// ---- SelfTests/TestCases/TestSuite_EventDelivery/Test_EventDeleteLostSequence.TcPOU
{region 'Documentation'}
(*!
<summary>Verifies deletion progress stops at retained events when the requested sequence was lost.</summary>
<description>
Four primary events plus the capacity diagnostic fill five usable slots. Publications 6
and 7 fail, creating a real sequence gap. Request 6 exhausts the retained prefix at 5 and
appends diagnostic 8. Request 7 must leave that newer head intact and append diagnostic 9.
No sequence, FIFO index or private subject field is modified to arrange these cases.
The real subject binds only local storage; expected findings remain in that storage.
Checking Assertions retain the outer selftest publisher. Each run reinitializes the subject.
</description>
*)
{endregion}
FUNCTION_BLOCK Test_EventDeleteLostSequence EXTENDS TestCaseBase
VAR
    FSubject : EventBuffer;
    FEvents : ARRAY[1..BufferLength] OF ST_Event;
    FFifo : ST_FifoStatus;
    FBufferStatus : ST_EventBufferStatus;
    FPerformed : BOOL;
    FChecked : BOOL;
    FLostTargets : AssertTrue;
    FLostTargetsMatches : BOOL;
    FActualProgress : AssertTrue;
    FActualProgressMatches : BOOL;
    FExhaustionDiagnostic : AssertTrue;
    FExhaustionDiagnosticMatches : BOOL;
    FNewerHeadPreserved : AssertTrue;
    FNewerHeadPreservedMatches : BOOL;
    FGapDiagnostic : AssertTrue;
    FGapDiagnosticMatches : BOOL;
END_VAR
VAR CONSTANT
    BufferLength : UINT := 6;
END_VAR

SUPER^();

{region 'Documentation'}
(*!
<summary>Contributes each checking Assertion once.</summary>
*)
{endregion}
METHOD PROTECTED AggregateResults
VAR_INPUT
    Aggregator : I_ResultAggregator; //! Borrowed result sink owned by the outer Test Case; add this test's checking Assertions without resetting or retaining the sink.
END_VAR
Aggregator.AddProvider(Provider := FLostTargets);
Aggregator.AddProvider(Provider := FActualProgress);
Aggregator.AddProvider(Provider := FExhaustionDiagnostic);
Aggregator.AddProvider(Provider := FNewerHeadPreserved);
Aggregator.AddProvider(Provider := FGapDiagnostic);
END_METHOD

{region 'Documentation'}
(*!
<summary>Requires all checking Assertions to be initialized.</summary>
*)
{endregion}
METHOD PROTECTED CheckInitialization : BOOL //! TRUE when the inherited initialization check and this concrete fixture check both accept the setup.
CheckInitialization := FALSE;
IF NOT SUPER^.CheckInitialization() THEN
    RETURN;
END_IF;

CheckInitialization := FLostTargets.IsInitialized
    AND FActualProgress.IsInitialized
    AND FExhaustionDiagnostic.IsInitialized
    AND FNewerHeadPreserved.IsInitialized
    AND FGapDiagnostic.IsInitialized;
END_METHOD

{region 'Documentation'}
(*!
<summary>Initializes the checking Assertions for one test state.</summary>
*)
{endregion}
METHOD PROTECTED Configure
FPreparationStateCount := 0;
FTestStateCount := 1;
FLostTargets.Initialize(Parent := THIS^,
    AssertionName := 'LostTargets');
FActualProgress.Initialize(Parent := THIS^,
    AssertionName := 'ActualProgress');
FExhaustionDiagnostic.Initialize(Parent := THIS^,
    AssertionName := 'ExhaustionDiagnostic');
FNewerHeadPreserved.Initialize(Parent := THIS^,
    AssertionName := 'NewerHeadPreserved');
FGapDiagnostic.Initialize(Parent := THIS^,
    AssertionName := 'GapDiagnostic');
END_METHOD

{region 'Documentation'}
(*!
<summary>Fills the buffer and verifies that sequences 6 and 7 were assigned but not retained.</summary>
*)
{endregion}
METHOD PRIVATE CreateLostTargets
VAR
    Index : UINT;
    WriteResult : INT;
END_VAR
FLostTargetsMatches := TRUE;
FOR Index := 1 TO 4 DO
    WriteResult := FSubject.PublishEvent(Event := CreateFrameworkEvent(Name := 'LocalGap',
        State := E_State.Running,
        Severity := E_EventSeverity.Info,
        Message := UINT_TO_STRING(Index)));
    FLostTargetsMatches := FLostTargetsMatches AND (WriteResult = UINT_TO_INT(Index));
END_FOR;
FOR Index := 6 TO 7 DO
    WriteResult := FSubject.PublishEvent(Event := CreateFrameworkEvent(Name := 'Lost',
        State := E_State.Running,
        Severity := E_EventSeverity.Info,
        Message := UINT_TO_STRING(Index)));
    FLostTargetsMatches := FLostTargetsMatches AND (WriteResult = TO_INT(E_FifoResult.NoTransfer));
END_FOR;
FLostTargetsMatches := FLostTargetsMatches AND FFifo.BufferFull
    AND (FFifo.ElementCount = 5) AND (FFifo.IndexOut = 1) AND (FFifo.IndexIn = 6)
    AND (FBufferStatus.SequenceId = 7) AND (FBufferStatus.DeletedSequenceId = 0)
    AND (FBufferStatus.LostEventCount = 2);
FOR Index := 1 TO 5 DO
    FLostTargetsMatches := FLostTargetsMatches AND (FEvents[Index].SequenceId = UINT_TO_UDINT(Index));
END_FOR;
END_METHOD

{region 'Documentation'}
(*!
<summary>A lost target below the current head must not delete that newer event or advance the watermark.</summary>
*)
{endregion}
METHOD PRIVATE DeleteBeforeNewerHead
VAR
    Request : UDINT;
    HeadBeforeRequest : ST_Event;
END_VAR
HeadBeforeRequest := FEvents[6];
Request := 7;
FSubject.ProcessDeleteRequest(SequenceId := Request);
FNewerHeadPreservedMatches := (Request = 0) AND (FBufferStatus.DeletedSequenceId = 5)
    AND (FBufferStatus.LostEventCount = 2)
    AND (FFifo.IndexOut = 6) AND (FFifo.IndexIn = 2) AND (FFifo.ElementCount = 2)
    AND (FEvents[6].SequenceId = 8)
    AND (FEvents[6].SequenceId = HeadBeforeRequest.SequenceId)
    AND (FEvents[6].Timestamp = HeadBeforeRequest.Timestamp)
    AND (FEvents[6].OwnerScope = HeadBeforeRequest.OwnerScope)
    AND (FEvents[6].EventType = HeadBeforeRequest.EventType)
    AND (FEvents[6].Severity = HeadBeforeRequest.Severity)
    AND (FEvents[6].Name = HeadBeforeRequest.Name)
    AND (FEvents[6].ResourceName = HeadBeforeRequest.ResourceName)
    AND (FEvents[6].State = HeadBeforeRequest.State)
    AND (FEvents[6].Result = HeadBeforeRequest.Result)
    AND (FEvents[6].Message = HeadBeforeRequest.Message);
FGapDiagnosticMatches := (FBufferStatus.SequenceId = 9)
    AND (FEvents[1].SequenceId = 9) AND (FEvents[1].OwnerScope = E_OwnerScope.Framework)
    AND (FEvents[1].EventType = E_EventType.Framework)
    AND (FEvents[1].Severity = E_EventSeverity.Warning) AND (FEvents[1].Name = 'EventBuffer');
END_METHOD

{region 'Documentation'}
(*!
<summary>Deletion exhausts at sequence 5; the newly appended diagnostic is not part of that prefix.</summary>
*)
{endregion}
METHOD PRIVATE DeleteBeyondRetainedTail
VAR
    Request : UDINT;
    Index : UINT;
END_VAR
Request := 6;
FSubject.ProcessDeleteRequest(SequenceId := Request);
FActualProgressMatches := (Request = 0) AND (FBufferStatus.DeletedSequenceId = 5)
    AND (FBufferStatus.LostEventCount = 2);
FOR Index := 1 TO 5 DO
    FActualProgressMatches := FActualProgressMatches AND (FEvents[Index].SequenceId = 0)
        AND (FEvents[Index].Timestamp = 0) AND (FEvents[Index].Name = '') AND (FEvents[Index].Message = '');
END_FOR;
FExhaustionDiagnosticMatches := (FBufferStatus.SequenceId = 8)
    AND NOT FFifo.BufferEmpty AND (FFifo.ElementCount = 1)
    AND (FFifo.IndexOut = 6) AND (FFifo.IndexIn = 1)
    AND (FEvents[6].SequenceId = 8) AND (FEvents[6].OwnerScope = E_OwnerScope.Framework)
    AND (FEvents[6].EventType = E_EventType.Framework)
    AND (FEvents[6].Severity = E_EventSeverity.Warning) AND (FEvents[6].Name = 'EventBuffer');
END_METHOD

{region 'Documentation'}
(*!
<summary>Creates two lost targets through overflow, then exercises exhaustion and a newer FIFO head.</summary>
*)
{endregion}
METHOD PRIVATE ExerciseBuffer
IF NOT FSubject.Initialize(Buffer := FEvents,
    FifoControl := FFifo,
    Status := FBufferStatus) THEN
    Error(Message := 'Local Event Buffer initialization failed.');
    RETURN;
END_IF;

CreateLostTargets();
DeleteBeyondRetainedTail();
DeleteBeforeNewerHead();
END_METHOD

{region 'Documentation'}
(*!
<summary>Completes abort without asynchronous work.</summary>
*)
{endregion}
METHOD PROTECTED ProcessAbort
VAR_INPUT
    Enable : BOOL; //! Phase permission supplied by the owning Test Case; FALSE does not authorize progression, while observation may continue.
END_VAR
IF Enable THEN
    CompleteAbort();
END_IF;
END_METHOD

{region 'Documentation'}
(*!
<summary>Evaluates captured observations after the scenario has finished.</summary>
*)
{endregion}
METHOD PROTECTED ProcessAssertions
VAR_INPUT
    Enable : BOOL; //! Phase permission supplied by the owning Test Case; FALSE does not authorize progression, while observation may continue.
END_VAR
VAR
    Evaluate : BOOL;
END_VAR
Evaluate := Enable AND FPerformed;
FLostTargets(Enable := Evaluate,
    State := State,
    IN := FLostTargetsMatches);
FActualProgress(Enable := Evaluate,
    State := State,
    IN := FActualProgressMatches);
FExhaustionDiagnostic(Enable := Evaluate,
    State := State,
    IN := FExhaustionDiagnosticMatches);
FNewerHeadPreserved(Enable := Evaluate,
    State := State,
    IN := FNewerHeadPreservedMatches);
FGapDiagnostic(Enable := Evaluate,
    State := State,
    IN := FGapDiagnosticMatches);
IF Evaluate THEN
    FChecked := TRUE;
END_IF;
END_METHOD

{region 'Documentation'}
(*!
<summary>No Preparation phase is needed.</summary>
*)
{endregion}
METHOD PROTECTED ProcessPreparations
VAR_INPUT
    // SA0033: Required override without Preparation work.
    {attribute 'analysis' := '-33'}
    Enable : BOOL; //! Phase permission supplied by the owning Test Case; FALSE does not authorize progression, while observation may continue.
END_VAR
END_METHOD

{region 'Documentation'}
(*!
<summary>Resets observations and schedules a fresh subject initialization.</summary>
*)
{endregion}
METHOD PROTECTED ProcessReset
FPerformed := FALSE;
FChecked := FALSE;
FLostTargets.Reset();
FLostTargetsMatches := FALSE;
FActualProgress.Reset();
FActualProgressMatches := FALSE;
FExhaustionDiagnostic.Reset();
FExhaustionDiagnosticMatches := FALSE;
FNewerHeadPreserved.Reset();
FNewerHeadPreservedMatches := FALSE;
FGapDiagnostic.Reset();
FGapDiagnosticMatches := FALSE;
CompleteReset();
END_METHOD

{region 'Documentation'}
(*!
<summary>Runs the bounded scenario once before Assertion evaluation.</summary>
*)
{endregion}
METHOD PROTECTED ProcessTests
VAR_INPUT
    Enable : BOOL; //! Phase permission supplied by the owning Test Case; FALSE does not authorize progression, while observation may continue.
END_VAR
IF NOT Enable THEN
    RETURN;
END_IF;
IF FChecked THEN
    CompleteTests();
    RETURN;
END_IF;

IF NOT FPerformed THEN
    ExerciseBuffer();
    FPerformed := TRUE;
END_IF;
END_METHOD

END_FUNCTION_BLOCK

// ---- SelfTests/TestCases/TestSuite_EventDelivery/Test_EventDeleteCommandBoundary.TcPOU
{region 'Documentation'}
(*!
<summary>Verifies DeleteSequenceId consumption at explicit call boundaries across successive PLC cycles.</summary>
<description>
Uses the actual field of a local ST_EventBufferCommand as VAR_IN_OUT, not a copied request.
A higher watermark replaces an earlier value before the call. Another is queued after return,
survives publication in the next cycle and is consumed only by the following delete call.
Zero after successful or rejected processing must not replay deletion or diagnostics.
No write occurs inside ProcessDeleteRequest: this scenario does not exercise its changed-value
branch or establish atomicity against ADS writes between comparison and clearing.
The real subject binds only local storage; expected findings remain in that storage.
Checking Assertions retain the outer selftest publisher. Each run reinitializes the subject.
</description>
*)
{endregion}
FUNCTION_BLOCK Test_EventDeleteCommandBoundary EXTENDS TestCaseBase
VAR
    FSubject : EventBuffer;
    FEvents : ARRAY[1..BufferLength] OF ST_Event;
    FFifo : ST_FifoStatus;
    FBufferStatus : ST_EventBufferStatus;
    FPerformed : BOOL;
    FChecked : BOOL;
    FCommands : ST_EventBufferCommand;
    FStep : UINT;
    FBeforeCall : AssertTrue;
    FBeforeCallMatches : BOOL;
    FPending : AssertTrue;
    FPendingMatches : BOOL;
    FNextCall : AssertTrue;
    FNextCallMatches : BOOL;
    FZeroNoReplay : AssertTrue;
    FZeroNoReplayMatches : BOOL;
    FRejectedNoReplay : AssertTrue;
    FRejectedNoReplayMatches : BOOL;
END_VAR
VAR CONSTANT
    BufferLength : UINT := 10;
    Arrange : UINT := 0;
    ReplaceBeforeCall : UINT := 1;
    ObservePending : UINT := 2;
    ConsumePending : UINT := 3;
    ObserveCleared : UINT := 4;
    RejectFuture : UINT := 5;
    ObserveRejected : UINT := 6;
END_VAR

SUPER^();

{region 'Documentation'}
(*!
<summary>Contributes each checking Assertion once.</summary>
*)
{endregion}
METHOD PROTECTED AggregateResults
VAR_INPUT
    Aggregator : I_ResultAggregator; //! Borrowed result sink owned by the outer Test Case; add this test's checking Assertions without resetting or retaining the sink.
END_VAR
Aggregator.AddProvider(Provider := FBeforeCall);
Aggregator.AddProvider(Provider := FPending);
Aggregator.AddProvider(Provider := FNextCall);
Aggregator.AddProvider(Provider := FZeroNoReplay);
Aggregator.AddProvider(Provider := FRejectedNoReplay);
END_METHOD

{region 'Documentation'}
(*!
<summary>Requires all checking Assertions to be initialized.</summary>
*)
{endregion}
METHOD PROTECTED CheckInitialization : BOOL //! TRUE when the inherited initialization check and this concrete fixture check both accept the setup.
CheckInitialization := FALSE;
IF NOT SUPER^.CheckInitialization() THEN
    RETURN;
END_IF;

CheckInitialization := FBeforeCall.IsInitialized
    AND FPending.IsInitialized
    AND FNextCall.IsInitialized
    AND FZeroNoReplay.IsInitialized
    AND FRejectedNoReplay.IsInitialized;
END_METHOD

{region 'Documentation'}
(*!
<summary>Initializes the checking Assertions for one test state.</summary>
*)
{endregion}
METHOD PROTECTED Configure
FPreparationStateCount := 0;
FTestStateCount := 1;
FBeforeCall.Initialize(Parent := THIS^,
    AssertionName := 'BeforeCall');
FPending.Initialize(Parent := THIS^,
    AssertionName := 'Pending');
FNextCall.Initialize(Parent := THIS^,
    AssertionName := 'NextCall');
FZeroNoReplay.Initialize(Parent := THIS^,
    AssertionName := 'ZeroNoReplay');
FRejectedNoReplay.Initialize(Parent := THIS^,
    AssertionName := 'RejectedNoReplay');
END_METHOD

{region 'Documentation'}
(*!
<summary>Completes abort without asynchronous work.</summary>
*)
{endregion}
METHOD PROTECTED ProcessAbort
VAR_INPUT
    Enable : BOOL; //! Phase permission supplied by the owning Test Case; FALSE does not authorize progression, while observation may continue.
END_VAR
IF Enable THEN
    CompleteAbort();
END_IF;
END_METHOD

{region 'Documentation'}
(*!
<summary>Evaluates captured observations after the scenario has finished.</summary>
*)
{endregion}
METHOD PROTECTED ProcessAssertions
VAR_INPUT
    Enable : BOOL; //! Phase permission supplied by the owning Test Case; FALSE does not authorize progression, while observation may continue.
END_VAR
VAR
    Evaluate : BOOL;
END_VAR
Evaluate := Enable AND FPerformed;
FBeforeCall(Enable := Evaluate,
    State := State,
    IN := FBeforeCallMatches);
FPending(Enable := Evaluate,
    State := State,
    IN := FPendingMatches);
FNextCall(Enable := Evaluate,
    State := State,
    IN := FNextCallMatches);
FZeroNoReplay(Enable := Evaluate,
    State := State,
    IN := FZeroNoReplayMatches);
FRejectedNoReplay(Enable := Evaluate,
    State := State,
    IN := FRejectedNoReplayMatches);
IF Evaluate THEN
    FChecked := TRUE;
END_IF;
END_METHOD

{region 'Documentation'}
(*!
<summary>No Preparation phase is needed.</summary>
*)
{endregion}
METHOD PROTECTED ProcessPreparations
VAR_INPUT
    // SA0033: Required override without Preparation work.
    {attribute 'analysis' := '-33'}
    Enable : BOOL; //! Phase permission supplied by the owning Test Case; FALSE does not authorize progression, while observation may continue.
END_VAR
END_METHOD

{region 'Documentation'}
(*!
<summary>Resets observations and schedules a fresh subject initialization.</summary>
*)
{endregion}
METHOD PROTECTED ProcessReset
FPerformed := FALSE;
FChecked := FALSE;
FStep := Arrange;
FCommands.Reset := FALSE;
FCommands.DeleteSequenceId := 0;
FBeforeCall.Reset();
FBeforeCallMatches := FALSE;
FPending.Reset();
FPendingMatches := FALSE;
FNextCall.Reset();
FNextCallMatches := FALSE;
FZeroNoReplay.Reset();
FZeroNoReplayMatches := FALSE;
FRejectedNoReplay.Reset();
FRejectedNoReplayMatches := FALSE;
CompleteReset();
END_METHOD

{region 'Documentation'}
(*!
<summary>Advances the scenario until its final observation has been evaluated.</summary>
*)
{endregion}
METHOD PROTECTED ProcessTests
VAR_INPUT
    Enable : BOOL; //! Phase permission supplied by the owning Test Case; FALSE does not authorize progression, while observation may continue.
END_VAR
IF NOT Enable THEN
    RETURN;
END_IF;
IF FChecked THEN
    CompleteTests();
    RETURN;
END_IF;

IF NOT FPerformed THEN
    StateMachine();
END_IF;
END_METHOD

{region 'Documentation'}
(*!
<summary>Advances one boundary scenario step per enabled test cycle.</summary>
*)
{endregion}
METHOD PRIVATE StateMachine
VAR
    Index : UINT;
    WriteResult : INT;
END_VAR
CASE FStep OF
    Arrange:
        IF NOT FSubject.Initialize(Buffer := FEvents,
            FifoControl := FFifo,
            Status := FBufferStatus) THEN
            Error(Message := 'Local Event Buffer initialization failed.');
            RETURN;
        END_IF;
        FBeforeCallMatches := TRUE;
        FOR Index := 1 TO 4 DO
            WriteResult := FSubject.PublishEvent(Event := CreateFrameworkEvent(Name := 'LocalCommand',
                State := E_State.Running,
                Severity := E_EventSeverity.Info,
                Message := UINT_TO_STRING(Index)));
            FBeforeCallMatches := FBeforeCallMatches AND (WriteResult = UINT_TO_INT(Index));
        END_FOR;
        FStep := ReplaceBeforeCall;

    ReplaceBeforeCall:
        FCommands.DeleteSequenceId := 1;
        FCommands.DeleteSequenceId := 2;
        FSubject.ProcessDeleteRequest(SequenceId := FCommands.DeleteSequenceId);
        FBeforeCallMatches := FBeforeCallMatches AND (FCommands.DeleteSequenceId = 0)
            AND (FBufferStatus.DeletedSequenceId = 2) AND (FBufferStatus.SequenceId = 4)
            AND (FFifo.IndexOut = 3) AND (FFifo.IndexIn = 5) AND (FFifo.ElementCount = 2)
            AND (FEvents[1].SequenceId = 0) AND (FEvents[2].SequenceId = 0)
            AND (FEvents[3].SequenceId = 3) AND (FEvents[4].SequenceId = 4);
        FCommands.DeleteSequenceId := 4;
        FStep := ObservePending;

    ObservePending:
        WriteResult := FSubject.PublishEvent(Event := CreateFrameworkEvent(Name := 'LocalCommand',
            State := E_State.Running,
            Severity := E_EventSeverity.Info,
            Message := 'Published while deletion is pending.'));
        FPendingMatches := (WriteResult = 5) AND (FCommands.DeleteSequenceId = 4)
            AND (FBufferStatus.DeletedSequenceId = 2) AND (FBufferStatus.SequenceId = 5)
            AND (FFifo.IndexOut = 3) AND (FFifo.IndexIn = 6) AND (FFifo.ElementCount = 3)
            AND (FEvents[3].SequenceId = 3) AND (FEvents[4].SequenceId = 4)
            AND (FEvents[5].SequenceId = 5);
        FStep := ConsumePending;

    ConsumePending:
        FSubject.ProcessDeleteRequest(SequenceId := FCommands.DeleteSequenceId);
        FNextCallMatches := (FCommands.DeleteSequenceId = 0)
            AND (FBufferStatus.DeletedSequenceId = 4) AND (FBufferStatus.SequenceId = 5)
            AND (FFifo.IndexOut = 5) AND (FFifo.IndexIn = 6) AND (FFifo.ElementCount = 1)
            AND (FEvents[3].SequenceId = 0) AND (FEvents[4].SequenceId = 0)
            AND (FEvents[5].SequenceId = 5);
        FStep := ObserveCleared;

    ObserveCleared:
        FSubject.ProcessDeleteRequest(SequenceId := FCommands.DeleteSequenceId);
        FZeroNoReplayMatches := (FCommands.DeleteSequenceId = 0)
            AND (FBufferStatus.DeletedSequenceId = 4) AND (FBufferStatus.SequenceId = 5)
            AND (FFifo.IndexOut = 5) AND (FFifo.IndexIn = 6) AND (FFifo.ElementCount = 1)
            AND (FEvents[5].SequenceId = 5) AND (FBufferStatus.LostEventCount = 0);
        FCommands.DeleteSequenceId := 100;
        FStep := RejectFuture;

    RejectFuture:
        FSubject.ProcessDeleteRequest(SequenceId := FCommands.DeleteSequenceId);
        FRejectedNoReplayMatches := (FCommands.DeleteSequenceId = 0)
            AND (FBufferStatus.DeletedSequenceId = 4) AND (FBufferStatus.SequenceId = 6)
            AND (FFifo.IndexOut = 5) AND (FFifo.IndexIn = 7) AND (FFifo.ElementCount = 2)
            AND (FEvents[5].SequenceId = 5)
            AND (FEvents[6].SequenceId = 6) AND (FEvents[6].Name = 'EventBuffer')
            AND (FEvents[6].EventType = E_EventType.Framework)
            AND (FEvents[6].Severity = E_EventSeverity.Warning);
        FStep := ObserveRejected;

    ObserveRejected:
        FSubject.ProcessDeleteRequest(SequenceId := FCommands.DeleteSequenceId);
        FRejectedNoReplayMatches := FRejectedNoReplayMatches AND (FCommands.DeleteSequenceId = 0)
            AND (FBufferStatus.DeletedSequenceId = 4) AND (FBufferStatus.SequenceId = 6)
            AND (FFifo.IndexOut = 5) AND (FFifo.IndexIn = 7) AND (FFifo.ElementCount = 2)
            AND (FEvents[5].SequenceId = 5) AND (FEvents[6].SequenceId = 6)
            AND (FBufferStatus.LostEventCount = 0);
        FPerformed := TRUE;

ELSE
    Error(Message := 'Unknown delete-command test step.');
END_CASE;
END_METHOD

END_FUNCTION_BLOCK

// ---- SelfTests/TestSuites/TestSuite_EventReservation.TcPOU
{region 'Documentation'}
(*!
<summary>Groups real event reservation, admission and hierarchical release tests on isolated storage.</summary>
*)
{endregion}
FUNCTION_BLOCK TestSuite_EventReservation EXTENDS TestSuiteBase
VAR
    FSubjectParent : I_RunControl;
    FResetAccounting : Test_ResetReservationAccounting;
    FExecutionAccounting : Test_ExecutionReservationAccounting;
    FAdmission : Test_ReservationAdmission;
    FImpossibleReset : Test_ImpossibleResetBudget;
    FImpossibleExecution : Test_ImpossibleExecutionBudget;
    FActiveReservationLoss : Test_ActiveReservationLoss;
    FHierarchicalRelease : Test_HierarchicalReservationRelease;
    FLateResetRelease : Test_LateResetReservationRelease;
    FTestCases : ARRAY[1..TestCaseCapacity] OF I_TestCase;
END_VAR
VAR CONSTANT
    TestCaseCapacity : UINT := 8;
END_VAR

SUPER^();

{region 'Documentation'}
(*!
<summary>Supplies the existing root identity to isolated Suite subjects before initialization.</summary>
*)
{endregion}
METHOD PUBLIC BindSubjectParent
VAR_INPUT
    Parent : I_RunControl; //! Borrowed identity parent retained for isolated subject initialization; keep the Run-Control alive through subject use.
END_VAR
FSubjectParent := Parent;
END_METHOD

{region 'Documentation'}
(*!
<summary>Initializes and registers the isolated event scenarios for serial execution.</summary>
*)
{endregion}
METHOD PROTECTED Configure
VAR_IN_OUT
    // SA0167: Borrowed owner builder; no temporary instance is created.
    {attribute 'analysis' := '-167'}
    Builder : TestSuiteConfigurationBuilder; //! Borrowed owner configuration builder used only during this Configure call; register this owner's concrete children.
END_VAR
VAR
    TestConfig : ST_TestCaseConfig;
END_VAR
Builder.Initialize(Mode := E_OrchestrationMode.Serial,
    TestCases := FTestCases);
FResetAccounting.Initialize(Parent := THIS^,
    TestName := 'ResetAccounting',
    Config := TestConfig);
Builder.Register(TestCase := FResetAccounting);

FExecutionAccounting.Initialize(Parent := THIS^,
    TestName := 'ExecutionAccounting',
    Config := TestConfig);
Builder.Register(TestCase := FExecutionAccounting);

FAdmission.BindSubjectParent(Parent := THIS^);
FAdmission.Initialize(Parent := THIS^,
    TestName := 'Admission',
    Config := TestConfig);
Builder.Register(TestCase := FAdmission);

FImpossibleReset.BindSubjectParent(Parent := THIS^);
FImpossibleReset.Initialize(Parent := THIS^,
    TestName := 'ImpossibleReset',
    Config := TestConfig);
Builder.Register(TestCase := FImpossibleReset);

FImpossibleExecution.BindSubjectParent(Parent := THIS^);
FImpossibleExecution.Initialize(Parent := THIS^,
    TestName := 'ImpossibleExecution',
    Config := TestConfig);
Builder.Register(TestCase := FImpossibleExecution);

FActiveReservationLoss.BindSubjectParent(Parent := THIS^);
FActiveReservationLoss.Initialize(Parent := THIS^,
    TestName := 'ActiveReservationLoss',
    Config := TestConfig);
Builder.Register(TestCase := FActiveReservationLoss);

FHierarchicalRelease.BindSubjectParent(Parent := FSubjectParent);
FHierarchicalRelease.Initialize(Parent := THIS^,
    TestName := 'HierarchicalRelease',
    Config := TestConfig);
Builder.Register(TestCase := FHierarchicalRelease);

FLateResetRelease.BindSubjectParent(Parent := FSubjectParent);
FLateResetRelease.Initialize(Parent := THIS^,
    TestName := 'LateResetRelease',
    Config := TestConfig);
Builder.Register(TestCase := FLateResetRelease);
END_METHOD

{region 'Documentation'}
(*!
<summary>Returns a registered scenario using its original array index.</summary>
*)
{endregion}
METHOD PUBLIC GetTestCase : I_TestCase //! Typed child interface at the original array index; zero when no entry is available.
VAR_INPUT
    Index : DINT; //! Original occupied child-array index, rather than an ordinal position.
END_VAR
GetTestCase := 0;
IF (ChildCount = 0) OR (Index < ChildArrayLowerBound)
    OR (DINT_TO_LINT(Index) >= DINT_TO_LINT(ChildArrayLowerBound) + UINT_TO_LINT(ChildCount)) THEN
    RETURN;
END_IF;
GetTestCase := FTestCases[Index];
END_METHOD

{region 'Documentation'}
(*!
<summary>Calls each owned scenario once per initialized Suite cycle.</summary>
*)
{endregion}
METHOD PROTECTED ProcessTestCases
FResetAccounting();
FExecutionAccounting();
FAdmission();
FImpossibleReset();
FImpossibleExecution();
FActiveReservationLoss();
FHierarchicalRelease();
FLateResetRelease();
END_METHOD

END_FUNCTION_BLOCK

// ---- SelfTests/TestCases/TestSuite_EventReservation/Test_ResetReservationAccounting.TcPOU
{region 'Documentation'}
(*!
<summary>Checks reset reservation accounting on an exactly sized local Event Buffer.</summary>
<description>
Local counters represent two independent reservation callers, not child FB instances.
The budget is four Suite plus three Test Case entries and one shared Reset headroom.
Storage includes the FIFO spare position. These API tests do not prove owner admission.
Owner budget calculation and child dispatch are checked by separate integration scenarios.
The real subject binds only local storage; expected findings remain in that storage.
Checking Assertions retain the outer selftest publisher. Each run reinitializes the subject.
</description>
*)
{endregion}
FUNCTION_BLOCK Test_ResetReservationAccounting EXTENDS TestCaseBase
VAR
    FSubject : EventBuffer;
    FEvents : ARRAY[1..BufferLength] OF ST_Event;
    FFifo : ST_FifoStatus;
    FBufferStatus : ST_EventBufferStatus;
    FPerformed : BOOL;
    FChecked : BOOL;
    FSuiteReserved : UINT;
    FChildReserved : UINT;
    FInitialFifo : ST_FifoStatus;
    FBinding : AssertTrue;
    FBindingMatches : BOOL;
    FSuiteContribution : AssertTrue;
    FSuiteContributionMatches : BOOL;
    FCombinedContributions : AssertTrue;
    FCombinedContributionsMatches : BOOL;
    FRejectedReservation : AssertTrue;
    FRejectedReservationMatches : BOOL;
    FChildRelease : AssertTrue;
    FChildReleaseMatches : BOOL;
    FBalancedRelease : AssertTrue;
    FBalancedReleaseMatches : BOOL;
    FRepeatedRelease : AssertTrue;
    FRepeatedReleaseMatches : BOOL;
    FReadableDataUnchanged : AssertTrue;
    FReadableDataUnchangedMatches : BOOL;
END_VAR
VAR CONSTANT
    SuiteBudget : UINT := GVL_Constants.TestSuiteResetEventCount;
    ChildBudget : UINT := GVL_Constants.TestCaseResetEventCount;
    Headroom : UINT := Param_EventBuffer.EventBufferResetHeadroom;
    BufferLength : UINT := SuiteBudget + ChildBudget + Headroom + 1;
END_VAR

SUPER^();

{region 'Documentation'}
(*!
<summary>Contributes each checking Assertion once.</summary>
*)
{endregion}
METHOD PROTECTED AggregateResults
VAR_INPUT
    Aggregator : I_ResultAggregator; //! Borrowed result sink owned by the outer Test Case; add this test's checking Assertions without resetting or retaining the sink.
END_VAR
Aggregator.AddProvider(Provider := FBinding);
Aggregator.AddProvider(Provider := FSuiteContribution);
Aggregator.AddProvider(Provider := FCombinedContributions);
Aggregator.AddProvider(Provider := FRejectedReservation);
Aggregator.AddProvider(Provider := FChildRelease);
Aggregator.AddProvider(Provider := FBalancedRelease);
Aggregator.AddProvider(Provider := FRepeatedRelease);
Aggregator.AddProvider(Provider := FReadableDataUnchanged);
END_METHOD

{region 'Documentation'}
(*!
<summary>Requires all checking Assertions to be initialized.</summary>
*)
{endregion}
METHOD PROTECTED CheckInitialization : BOOL //! TRUE when the inherited initialization check and this concrete fixture check both accept the setup.
CheckInitialization := FALSE;
IF NOT SUPER^.CheckInitialization() THEN
    RETURN;
END_IF;

CheckInitialization := FBinding.IsInitialized
    AND FSuiteContribution.IsInitialized
    AND FCombinedContributions.IsInitialized
    AND FRejectedReservation.IsInitialized
    AND FChildRelease.IsInitialized
    AND FBalancedRelease.IsInitialized
    AND FRepeatedRelease.IsInitialized
    AND FReadableDataUnchanged.IsInitialized;
END_METHOD

{region 'Documentation'}
(*!
<summary>Initializes the checking Assertions for one test state.</summary>
*)
{endregion}
METHOD PROTECTED Configure
FPreparationStateCount := 0;
FTestStateCount := 1;
FBinding.Initialize(Parent := THIS^,
    AssertionName := 'Binding');
FSuiteContribution.Initialize(Parent := THIS^,
    AssertionName := 'SuiteContribution');
FCombinedContributions.Initialize(Parent := THIS^,
    AssertionName := 'CombinedContributions');
FRejectedReservation.Initialize(Parent := THIS^,
    AssertionName := 'RejectedReservation');
FChildRelease.Initialize(Parent := THIS^,
    AssertionName := 'ChildRelease');
FBalancedRelease.Initialize(Parent := THIS^,
    AssertionName := 'BalancedRelease');
FRepeatedRelease.Initialize(Parent := THIS^,
    AssertionName := 'RepeatedRelease');
FReadableDataUnchanged.Initialize(Parent := THIS^,
    AssertionName := 'ReadableDataUnchanged');
END_METHOD

{region 'Documentation'}
(*!
<summary>Checks local contributions and buffer-wide accounting at exact capacity.</summary>
*)
{endregion}
METHOD PRIVATE ExerciseBuffer
VAR
    Initialized : BOOL;
END_VAR
FSuiteReserved := 0;
FChildReserved := 0;
Initialized := FSubject.Initialize(Buffer := FEvents,
    FifoControl := FFifo,
    Status := FBufferStatus);
FBindingMatches := Initialized
    AND (FSubject.Capacity = BufferLength - 1)
    AND (FSubject.FreeEntryCount = BufferLength - 1)
    AND (FSubject.ReservedEntryCount = 0);
IF NOT Initialized THEN
    RETURN;
END_IF;

FInitialFifo := FFifo;
ReserveBudgets();
RejectAdditionalReservation();
ReleaseBudgets();

FReadableDataUnchangedMatches := (FFifo.IndexIn = FInitialFifo.IndexIn)
    AND (FFifo.IndexOut = FInitialFifo.IndexOut)
    AND (FFifo.ElementCount = 0) AND FFifo.BufferEmpty
    AND (FSubject.FreeEntryCount = BufferLength - 1)
    AND (FBufferStatus.SequenceId = 0)
    AND (FBufferStatus.DeletedSequenceId = 0)
    AND (FBufferStatus.LostEventCount = 0);
END_METHOD

{region 'Documentation'}
(*!
<summary>Completes abort without asynchronous work.</summary>
*)
{endregion}
METHOD PROTECTED ProcessAbort
VAR_INPUT
    Enable : BOOL; //! Phase permission supplied by the owning Test Case; FALSE does not authorize progression, while observation may continue.
END_VAR
IF Enable THEN
    CompleteAbort();
END_IF;
END_METHOD

{region 'Documentation'}
(*!
<summary>Evaluates captured observations after the scenario has finished.</summary>
*)
{endregion}
METHOD PROTECTED ProcessAssertions
VAR_INPUT
    Enable : BOOL; //! Phase permission supplied by the owning Test Case; FALSE does not authorize progression, while observation may continue.
END_VAR
VAR
    Evaluate : BOOL;
END_VAR
Evaluate := Enable AND FPerformed;
FBinding(Enable := Evaluate,
    State := State,
    IN := FBindingMatches);
FSuiteContribution(Enable := Evaluate,
    State := State,
    IN := FSuiteContributionMatches);
FCombinedContributions(Enable := Evaluate,
    State := State,
    IN := FCombinedContributionsMatches);
FRejectedReservation(Enable := Evaluate,
    State := State,
    IN := FRejectedReservationMatches);
FChildRelease(Enable := Evaluate,
    State := State,
    IN := FChildReleaseMatches);
FBalancedRelease(Enable := Evaluate,
    State := State,
    IN := FBalancedReleaseMatches);
FRepeatedRelease(Enable := Evaluate,
    State := State,
    IN := FRepeatedReleaseMatches);
FReadableDataUnchanged(Enable := Evaluate,
    State := State,
    IN := FReadableDataUnchangedMatches);
IF Evaluate THEN
    FChecked := TRUE;
END_IF;
END_METHOD

{region 'Documentation'}
(*!
<summary>No Preparation phase is needed.</summary>
*)
{endregion}
METHOD PROTECTED ProcessPreparations
VAR_INPUT
    // SA0033: Required override without Preparation work.
    {attribute 'analysis' := '-33'}
    Enable : BOOL; //! Phase permission supplied by the owning Test Case; FALSE does not authorize progression, while observation may continue.
END_VAR
END_METHOD

{region 'Documentation'}
(*!
<summary>Resets observations and schedules a fresh subject initialization.</summary>
*)
{endregion}
METHOD PROTECTED ProcessReset
FPerformed := FALSE;
FChecked := FALSE;
FBinding.Reset();
FBindingMatches := FALSE;
FSuiteContribution.Reset();
FSuiteContributionMatches := FALSE;
FCombinedContributions.Reset();
FCombinedContributionsMatches := FALSE;
FRejectedReservation.Reset();
FRejectedReservationMatches := FALSE;
FChildRelease.Reset();
FChildReleaseMatches := FALSE;
FBalancedRelease.Reset();
FBalancedReleaseMatches := FALSE;
FRepeatedRelease.Reset();
FRepeatedReleaseMatches := FALSE;
FReadableDataUnchanged.Reset();
FReadableDataUnchangedMatches := FALSE;
CompleteReset();
END_METHOD

{region 'Documentation'}
(*!
<summary>Runs the bounded scenario once before Assertion evaluation.</summary>
*)
{endregion}
METHOD PROTECTED ProcessTests
VAR_INPUT
    Enable : BOOL; //! Phase permission supplied by the owning Test Case; FALSE does not authorize progression, while observation may continue.
END_VAR
IF NOT Enable THEN
    RETURN;
END_IF;
IF FChecked THEN
    CompleteTests();
    RETURN;
END_IF;

IF NOT FPerformed THEN
    ExerciseBuffer();
    FPerformed := TRUE;
END_IF;
END_METHOD

{region 'Documentation'}
(*!
<summary>Verifies rejection leaves both contributions and the aggregate unchanged.</summary>
*)
{endregion}
METHOD PRIVATE RejectAdditionalReservation
VAR
    Accepted : BOOL;
END_VAR
Accepted := FSubject.ReserveSpace(EntryCount := 1,
    HeadroomEntryCount := Headroom,
    OwnerReservedEntryCount := FChildReserved);
FRejectedReservationMatches := NOT Accepted
    AND (FSuiteReserved = SuiteBudget) AND (FChildReserved = ChildBudget)
    AND (FSubject.ReservedEntryCount = SuiteBudget + ChildBudget);
END_METHOD

{region 'Documentation'}
(*!
<summary>Releases each contribution independently and repeats an empty release.</summary>
*)
{endregion}
METHOD PRIVATE ReleaseBudgets
VAR
    Released : BOOL;
END_VAR
Released := FSubject.FreeReservedSpace(EntryCount := FChildReserved,
    OwnerReservedEntryCount := FChildReserved);
FChildReleaseMatches := Released
    AND (FChildReserved = 0) AND (FSuiteReserved = SuiteBudget)
    AND (FSubject.ReservedEntryCount = SuiteBudget);

Released := FSubject.FreeReservedSpace(EntryCount := FSuiteReserved,
    OwnerReservedEntryCount := FSuiteReserved);
FBalancedReleaseMatches := Released
    AND (FSuiteReserved = 0) AND (FChildReserved = 0)
    AND (FSubject.ReservedEntryCount = 0);

Released := FSubject.FreeReservedSpace(EntryCount := FChildReserved,
    OwnerReservedEntryCount := FChildReserved);
FRepeatedReleaseMatches := Released
    AND (FChildReserved = 0) AND (FSuiteReserved = 0)
    AND (FSubject.ReservedEntryCount = 0);
END_METHOD

{region 'Documentation'}
(*!
<summary>Reserves two independent contributions with shared headroom.</summary>
*)
{endregion}
METHOD PRIVATE ReserveBudgets
VAR
    Accepted : BOOL;
END_VAR
Accepted := FSubject.ReserveSpace(EntryCount := SuiteBudget,
    HeadroomEntryCount := Headroom,
    OwnerReservedEntryCount := FSuiteReserved);
FSuiteContributionMatches := Accepted
    AND (FSuiteReserved = SuiteBudget) AND (FChildReserved = 0)
    AND (FSubject.ReservedEntryCount = SuiteBudget);

Accepted := FSubject.ReserveSpace(EntryCount := ChildBudget,
    HeadroomEntryCount := Headroom,
    OwnerReservedEntryCount := FChildReserved);
FCombinedContributionsMatches := Accepted
    AND (FSuiteReserved = SuiteBudget) AND (FChildReserved = ChildBudget)
    AND (FSubject.ReservedEntryCount = SuiteBudget + ChildBudget)
    AND (FSubject.FreeEntryCount = FSubject.ReservedEntryCount + Headroom);
END_METHOD

END_FUNCTION_BLOCK

// ---- SelfTests/TestCases/TestSuite_EventReservation/Test_ExecutionReservationAccounting.TcPOU
{region 'Documentation'}
(*!
<summary>Checks execution reservation accounting on an exactly sized local Event Buffer.</summary>
<description>
Local counters represent two independent reservation callers, not child FB instances.
The budget is ten Suite entries plus eleven Test Case entries: zero Preparation states,
one test state, one Assertion and nine fixed lifecycle entries.
Storage includes the FIFO spare position. These API tests do not prove owner admission.
Owner budget calculation and child dispatch are checked by separate integration scenarios.
The real subject binds only local storage; expected findings remain in that storage.
Checking Assertions retain the outer selftest publisher. Each run reinitializes the subject.
</description>
*)
{endregion}
FUNCTION_BLOCK Test_ExecutionReservationAccounting EXTENDS TestCaseBase
VAR
    FSubject : EventBuffer;
    FEvents : ARRAY[1..BufferLength] OF ST_Event;
    FFifo : ST_FifoStatus;
    FBufferStatus : ST_EventBufferStatus;
    FPerformed : BOOL;
    FChecked : BOOL;
    FSuiteReserved : UINT;
    FChildReserved : UINT;
    FInitialFifo : ST_FifoStatus;
    FBinding : AssertTrue;
    FBindingMatches : BOOL;
    FSuiteContribution : AssertTrue;
    FSuiteContributionMatches : BOOL;
    FCombinedContributions : AssertTrue;
    FCombinedContributionsMatches : BOOL;
    FRejectedReservation : AssertTrue;
    FRejectedReservationMatches : BOOL;
    FChildRelease : AssertTrue;
    FChildReleaseMatches : BOOL;
    FBalancedRelease : AssertTrue;
    FBalancedReleaseMatches : BOOL;
    FRepeatedRelease : AssertTrue;
    FRepeatedReleaseMatches : BOOL;
    FReadableDataUnchanged : AssertTrue;
    FReadableDataUnchangedMatches : BOOL;
END_VAR
VAR CONSTANT
    SuiteBudget : UINT := GVL_Constants.TestSuiteExecutionEventCount;
    ChildBudget : UINT := 11;
    Headroom : UINT := Param_EventBuffer.EventBufferExecutionHeadroom;
    BufferLength : UINT := SuiteBudget + ChildBudget + Headroom + 1;
END_VAR

SUPER^();

{region 'Documentation'}
(*!
<summary>Contributes each checking Assertion once.</summary>
*)
{endregion}
METHOD PROTECTED AggregateResults
VAR_INPUT
    Aggregator : I_ResultAggregator; //! Borrowed result sink owned by the outer Test Case; add this test's checking Assertions without resetting or retaining the sink.
END_VAR
Aggregator.AddProvider(Provider := FBinding);
Aggregator.AddProvider(Provider := FSuiteContribution);
Aggregator.AddProvider(Provider := FCombinedContributions);
Aggregator.AddProvider(Provider := FRejectedReservation);
Aggregator.AddProvider(Provider := FChildRelease);
Aggregator.AddProvider(Provider := FBalancedRelease);
Aggregator.AddProvider(Provider := FRepeatedRelease);
Aggregator.AddProvider(Provider := FReadableDataUnchanged);
END_METHOD

{region 'Documentation'}
(*!
<summary>Requires all checking Assertions to be initialized.</summary>
*)
{endregion}
METHOD PROTECTED CheckInitialization : BOOL //! TRUE when the inherited initialization check and this concrete fixture check both accept the setup.
CheckInitialization := FALSE;
IF NOT SUPER^.CheckInitialization() THEN
    RETURN;
END_IF;

CheckInitialization := FBinding.IsInitialized
    AND FSuiteContribution.IsInitialized
    AND FCombinedContributions.IsInitialized
    AND FRejectedReservation.IsInitialized
    AND FChildRelease.IsInitialized
    AND FBalancedRelease.IsInitialized
    AND FRepeatedRelease.IsInitialized
    AND FReadableDataUnchanged.IsInitialized;
END_METHOD

{region 'Documentation'}
(*!
<summary>Initializes the checking Assertions for one test state.</summary>
*)
{endregion}
METHOD PROTECTED Configure
FPreparationStateCount := 0;
FTestStateCount := 1;
FBinding.Initialize(Parent := THIS^,
    AssertionName := 'Binding');
FSuiteContribution.Initialize(Parent := THIS^,
    AssertionName := 'SuiteContribution');
FCombinedContributions.Initialize(Parent := THIS^,
    AssertionName := 'CombinedContributions');
FRejectedReservation.Initialize(Parent := THIS^,
    AssertionName := 'RejectedReservation');
FChildRelease.Initialize(Parent := THIS^,
    AssertionName := 'ChildRelease');
FBalancedRelease.Initialize(Parent := THIS^,
    AssertionName := 'BalancedRelease');
FRepeatedRelease.Initialize(Parent := THIS^,
    AssertionName := 'RepeatedRelease');
FReadableDataUnchanged.Initialize(Parent := THIS^,
    AssertionName := 'ReadableDataUnchanged');
END_METHOD

{region 'Documentation'}
(*!
<summary>Checks local contributions and buffer-wide accounting at exact capacity.</summary>
*)
{endregion}
METHOD PRIVATE ExerciseBuffer
VAR
    Initialized : BOOL;
END_VAR
FSuiteReserved := 0;
FChildReserved := 0;
Initialized := FSubject.Initialize(Buffer := FEvents,
    FifoControl := FFifo,
    Status := FBufferStatus);
FBindingMatches := Initialized
    AND (FSubject.Capacity = BufferLength - 1)
    AND (FSubject.FreeEntryCount = BufferLength - 1)
    AND (FSubject.ReservedEntryCount = 0);
IF NOT Initialized THEN
    RETURN;
END_IF;

FInitialFifo := FFifo;
ReserveBudgets();
RejectAdditionalReservation();
ReleaseBudgets();

FReadableDataUnchangedMatches := (FFifo.IndexIn = FInitialFifo.IndexIn)
    AND (FFifo.IndexOut = FInitialFifo.IndexOut)
    AND (FFifo.ElementCount = 0) AND FFifo.BufferEmpty
    AND (FSubject.FreeEntryCount = BufferLength - 1)
    AND (FBufferStatus.SequenceId = 0)
    AND (FBufferStatus.DeletedSequenceId = 0)
    AND (FBufferStatus.LostEventCount = 0);
END_METHOD

{region 'Documentation'}
(*!
<summary>Completes abort without asynchronous work.</summary>
*)
{endregion}
METHOD PROTECTED ProcessAbort
VAR_INPUT
    Enable : BOOL; //! Phase permission supplied by the owning Test Case; FALSE does not authorize progression, while observation may continue.
END_VAR
IF Enable THEN
    CompleteAbort();
END_IF;
END_METHOD

{region 'Documentation'}
(*!
<summary>Evaluates captured observations after the scenario has finished.</summary>
*)
{endregion}
METHOD PROTECTED ProcessAssertions
VAR_INPUT
    Enable : BOOL; //! Phase permission supplied by the owning Test Case; FALSE does not authorize progression, while observation may continue.
END_VAR
VAR
    Evaluate : BOOL;
END_VAR
Evaluate := Enable AND FPerformed;
FBinding(Enable := Evaluate,
    State := State,
    IN := FBindingMatches);
FSuiteContribution(Enable := Evaluate,
    State := State,
    IN := FSuiteContributionMatches);
FCombinedContributions(Enable := Evaluate,
    State := State,
    IN := FCombinedContributionsMatches);
FRejectedReservation(Enable := Evaluate,
    State := State,
    IN := FRejectedReservationMatches);
FChildRelease(Enable := Evaluate,
    State := State,
    IN := FChildReleaseMatches);
FBalancedRelease(Enable := Evaluate,
    State := State,
    IN := FBalancedReleaseMatches);
FRepeatedRelease(Enable := Evaluate,
    State := State,
    IN := FRepeatedReleaseMatches);
FReadableDataUnchanged(Enable := Evaluate,
    State := State,
    IN := FReadableDataUnchangedMatches);
IF Evaluate THEN
    FChecked := TRUE;
END_IF;
END_METHOD

{region 'Documentation'}
(*!
<summary>No Preparation phase is needed.</summary>
*)
{endregion}
METHOD PROTECTED ProcessPreparations
VAR_INPUT
    // SA0033: Required override without Preparation work.
    {attribute 'analysis' := '-33'}
    Enable : BOOL; //! Phase permission supplied by the owning Test Case; FALSE does not authorize progression, while observation may continue.
END_VAR
END_METHOD

{region 'Documentation'}
(*!
<summary>Resets observations and schedules a fresh subject initialization.</summary>
*)
{endregion}
METHOD PROTECTED ProcessReset
FPerformed := FALSE;
FChecked := FALSE;
FBinding.Reset();
FBindingMatches := FALSE;
FSuiteContribution.Reset();
FSuiteContributionMatches := FALSE;
FCombinedContributions.Reset();
FCombinedContributionsMatches := FALSE;
FRejectedReservation.Reset();
FRejectedReservationMatches := FALSE;
FChildRelease.Reset();
FChildReleaseMatches := FALSE;
FBalancedRelease.Reset();
FBalancedReleaseMatches := FALSE;
FRepeatedRelease.Reset();
FRepeatedReleaseMatches := FALSE;
FReadableDataUnchanged.Reset();
FReadableDataUnchangedMatches := FALSE;
CompleteReset();
END_METHOD

{region 'Documentation'}
(*!
<summary>Runs the bounded scenario once before Assertion evaluation.</summary>
*)
{endregion}
METHOD PROTECTED ProcessTests
VAR_INPUT
    Enable : BOOL; //! Phase permission supplied by the owning Test Case; FALSE does not authorize progression, while observation may continue.
END_VAR
IF NOT Enable THEN
    RETURN;
END_IF;
IF FChecked THEN
    CompleteTests();
    RETURN;
END_IF;

IF NOT FPerformed THEN
    ExerciseBuffer();
    FPerformed := TRUE;
END_IF;
END_METHOD

{region 'Documentation'}
(*!
<summary>Verifies rejection leaves both contributions and the aggregate unchanged.</summary>
*)
{endregion}
METHOD PRIVATE RejectAdditionalReservation
VAR
    Accepted : BOOL;
END_VAR
Accepted := FSubject.ReserveSpace(EntryCount := 1,
    HeadroomEntryCount := Headroom,
    OwnerReservedEntryCount := FChildReserved);
FRejectedReservationMatches := NOT Accepted
    AND (FSuiteReserved = SuiteBudget) AND (FChildReserved = ChildBudget)
    AND (FSubject.ReservedEntryCount = SuiteBudget + ChildBudget);
END_METHOD

{region 'Documentation'}
(*!
<summary>Releases each contribution independently and repeats an empty release.</summary>
*)
{endregion}
METHOD PRIVATE ReleaseBudgets
VAR
    Released : BOOL;
END_VAR
Released := FSubject.FreeReservedSpace(EntryCount := FChildReserved,
    OwnerReservedEntryCount := FChildReserved);
FChildReleaseMatches := Released
    AND (FChildReserved = 0) AND (FSuiteReserved = SuiteBudget)
    AND (FSubject.ReservedEntryCount = SuiteBudget);

Released := FSubject.FreeReservedSpace(EntryCount := FSuiteReserved,
    OwnerReservedEntryCount := FSuiteReserved);
FBalancedReleaseMatches := Released
    AND (FSuiteReserved = 0) AND (FChildReserved = 0)
    AND (FSubject.ReservedEntryCount = 0);

Released := FSubject.FreeReservedSpace(EntryCount := FChildReserved,
    OwnerReservedEntryCount := FChildReserved);
FRepeatedReleaseMatches := Released
    AND (FChildReserved = 0) AND (FSuiteReserved = 0)
    AND (FSubject.ReservedEntryCount = 0);
END_METHOD

{region 'Documentation'}
(*!
<summary>Reserves two independent contributions with shared headroom.</summary>
*)
{endregion}
METHOD PRIVATE ReserveBudgets
VAR
    Accepted : BOOL;
END_VAR
Accepted := FSubject.ReserveSpace(EntryCount := SuiteBudget,
    HeadroomEntryCount := Headroom,
    OwnerReservedEntryCount := FSuiteReserved);
FSuiteContributionMatches := Accepted
    AND (FSuiteReserved = SuiteBudget) AND (FChildReserved = 0)
    AND (FSubject.ReservedEntryCount = SuiteBudget);

Accepted := FSubject.ReserveSpace(EntryCount := ChildBudget,
    HeadroomEntryCount := Headroom,
    OwnerReservedEntryCount := FChildReserved);
FCombinedContributionsMatches := Accepted
    AND (FSuiteReserved = SuiteBudget) AND (FChildReserved = ChildBudget)
    AND (FSubject.ReservedEntryCount = SuiteBudget + ChildBudget)
    AND (FSubject.FreeEntryCount = FSubject.ReservedEntryCount + Headroom);
END_METHOD

END_FUNCTION_BLOCK

// ---- SelfTests/TestCases/TestSuite_EventReservation/Test_ReservationAdmission.TcPOU
{region 'Documentation'}
(*!
<summary>Checks real Reset and Start admission before and after consumer deletion.</summary>
<description>

Isolation and call order

One real Orchestrator drives two real minimal Test Cases, called after the helper once per task cycle.
A thin child adapter observes held budgets at request entry; no scheduling or reservation response is simulated.
The collection double supplies fixed child interfaces. A local counter holds the concurrent Suite allowance;
Suite lifecycle and Suite budget calculation are not under test here.

Capacity pressure

Readable Info events reduce free capacity to one entry below admission. Three calls must remain silent
without a child request. Delete watermarks release occupancy, not reservations, and dispatch must resume.
Execution waiting must leave the children Idle and Ready. Completion is followed by three extra calls
to detect repeated dispatch. The outer Test Case timeout bounds unexpected non-completion.
The real subject binds only local storage; expected findings remain in that storage.
Checking Assertions retain the outer selftest publisher. Each run reinitializes the subject.
</description>
*)
{endregion}
FUNCTION_BLOCK Test_ReservationAdmission EXTENDS TestCaseBase
VAR
    FSubject : EventBuffer;
    FEvents : ARRAY[1..BufferLength] OF ST_Event;
    FFifo : ST_FifoStatus;
    FBufferStatus : ST_EventBufferStatus;
    FPerformed : BOOL;
    FChecked : BOOL;
    FSubjectParent : I_TestSuite;
    FOrchestrator : OrchestratorProbe;
    FCollection : OrchestrationCollectionDouble;
    FChildren : ARRAY[1..2] OF ReservationChildProbe;
    FChildViews : ARRAY[1..2] OF I_Orchestratable;
    FOwnerReserved : UINT;
    FStep : INT;
    FWaitCalls : UINT;
    FWaitingSequence : UDINT;
    FResetWaiting : AssertTrue;
    FResetWaitingMatches : BOOL;
    FExecutionWaiting : AssertTrue;
    FExecutionWaitingMatches : BOOL;
    FReservationBeforeRequest : AssertTrue;
    FReservationBeforeRequestMatches : BOOL;
    FSingleDispatch : AssertTrue;
    FSingleDispatchMatches : BOOL;
    FResumedExecution : AssertTrue;
    FResumedExecutionMatches : BOOL;
    FAccounting : AssertTrue;
    FAccountingMatches : BOOL;
    FConsumerRelease : AssertTrue;
    FConsumerReleaseMatches : BOOL;
    FStorageIntegrity : AssertTrue;
    FStorageIntegrityMatches : BOOL;
END_VAR
VAR CONSTANT
    BufferLength : UINT := 65;
    ChildExecutionBudget : UINT := 11;
    WaitingCalls : UINT := 3;
    Setup : INT := 0;
    WaitForResetCapacity : INT := 1;
    CompleteSubjectReset : INT := 2;
    PrepareExecution : INT := 3;
    WaitForExecutionCapacity : INT := 4;
    CompleteSubjectExecution : INT := 5;
    Finish : INT := 6;
END_VAR

SUPER^();

{region 'Documentation'}
(*!
<summary>Contributes each checking Assertion once.</summary>
*)
{endregion}
METHOD PROTECTED AggregateResults
VAR_INPUT
    Aggregator : I_ResultAggregator; //! Borrowed result sink owned by the outer Test Case; add this test's checking Assertions without resetting or retaining the sink.
END_VAR
Aggregator.AddProvider(Provider := FResetWaiting);
Aggregator.AddProvider(Provider := FExecutionWaiting);
Aggregator.AddProvider(Provider := FReservationBeforeRequest);
Aggregator.AddProvider(Provider := FSingleDispatch);
Aggregator.AddProvider(Provider := FResumedExecution);
Aggregator.AddProvider(Provider := FAccounting);
Aggregator.AddProvider(Provider := FConsumerRelease);
Aggregator.AddProvider(Provider := FStorageIntegrity);
END_METHOD

{region 'Documentation'}
(*!
<summary>Supplies child identity only; the actual outer Suite does not execute the isolated children.</summary>
*)
{endregion}
METHOD PUBLIC BindSubjectParent
VAR_INPUT
    Parent : I_TestSuite; //! Borrowed identity parent retained for isolated subject initialization; keep the Suite alive through subject use.
END_VAR
FSubjectParent := Parent;
END_METHOD

{region 'Documentation'}
(*!
<summary>Calls the real helper before real children once, then checks request and accounting evidence.</summary>
*)
{endregion}
METHOD PRIVATE CallSubject
VAR_INPUT
    Task : E_OrchestratorTask; //! Orchestration task assigned for this controlled subject call.
END_VAR
VAR
    Index : INT;
END_VAR
FOrchestrator(Task := Task);
FAccountingMatches := FAccountingMatches
    AND (FSubject.ReservedEntryCount = FOwnerReserved
        + FChildren[1].ReservedEntryCount + FChildren[2].ReservedEntryCount);
FOR Index := 1 TO 2 DO
    FReservationBeforeRequestMatches := FReservationBeforeRequestMatches
        AND FChildren[Index].RequestsReserved;
    FSingleDispatchMatches := FSingleDispatchMatches
        AND (FChildren[Index].ResetRequestCount <= 1)
        AND (FChildren[Index].StartRequestCount <= 1);
    FChildren[Index]();
END_FOR;
FStorageIntegrityMatches := FStorageIntegrityMatches
    AND NOT FFifo.ConfigError AND NOT FFifo.IndexError
    AND (FBufferStatus.LostEventCount = 0)
    AND NOT FCollection.InvalidAccess AND NOT FCollection.TraceOverflow;
IF FOrchestrator.Result = E_Result.Error THEN
    Error(Message := 'Reservation admission Orchestrator reported Error.');
END_IF;
END_METHOD

{region 'Documentation'}
(*!
<summary>Requires all checking Assertions to be initialized.</summary>
*)
{endregion}
METHOD PROTECTED CheckInitialization : BOOL //! TRUE when the inherited initialization check and this concrete fixture check both accept the setup.
CheckInitialization := FALSE;
IF NOT SUPER^.CheckInitialization() OR (FSubjectParent = 0) THEN
    RETURN;
END_IF;

CheckInitialization := FResetWaiting.IsInitialized
    AND FExecutionWaiting.IsInitialized
    AND FReservationBeforeRequest.IsInitialized
    AND FSingleDispatch.IsInitialized
    AND FResumedExecution.IsInitialized
    AND FAccounting.IsInitialized
    AND FConsumerRelease.IsInitialized
    AND FStorageIntegrity.IsInitialized;
END_METHOD

{region 'Documentation'}
(*!
<summary>Initializes the checking Assertions for one test state.</summary>
*)
{endregion}
METHOD PROTECTED Configure
FPreparationStateCount := 0;
FTestStateCount := 1;
FResetWaiting.Initialize(Parent := THIS^,
    AssertionName := 'ResetWaiting');
FExecutionWaiting.Initialize(Parent := THIS^,
    AssertionName := 'ExecutionWaiting');
FReservationBeforeRequest.Initialize(Parent := THIS^,
    AssertionName := 'ReservationBeforeRequest');
FSingleDispatch.Initialize(Parent := THIS^,
    AssertionName := 'SingleDispatch');
FResumedExecution.Initialize(Parent := THIS^,
    AssertionName := 'ResumedExecution');
FAccounting.Initialize(Parent := THIS^,
    AssertionName := 'Accounting');
FConsumerRelease.Initialize(Parent := THIS^,
    AssertionName := 'ConsumerRelease');
FStorageIntegrity.Initialize(Parent := THIS^,
    AssertionName := 'StorageIntegrity');
END_METHOD

{region 'Documentation'}
(*!
<summary>Uses the normal acknowledgement watermark without resetting reservations or sequence history.</summary>
*)
{endregion}
METHOD PRIVATE DeletePublishedEvents
VAR
    Watermark : UDINT;
    LastPublished : UDINT;
    ReservedBefore : UINT;
END_VAR
LastPublished := FBufferStatus.SequenceId;
Watermark := LastPublished;
ReservedBefore := FSubject.ReservedEntryCount;
FSubject.ProcessDeleteRequest(SequenceId := Watermark);
FConsumerReleaseMatches := FConsumerReleaseMatches
    AND (Watermark = 0) AND FFifo.BufferEmpty
    AND (FSubject.FreeEntryCount = FSubject.Capacity)
    AND (FBufferStatus.SequenceId = LastPublished)
    AND (FBufferStatus.DeletedSequenceId = LastPublished)
    AND (FSubject.ReservedEntryCount = ReservedBefore);
END_METHOD

{region 'Documentation'}
(*!
<summary>Creates real readable occupancy one entry short of child admission, with a bounded loop.</summary>
*)
{endregion}
METHOD PRIVATE FillToFreeCount
VAR_INPUT
    FreeCount : UINT; //! Target free-entry count reached by publishing bounded filler events; mismatch reports Error.
END_VAR
VAR
    Index : UINT;
    Filler : ST_Event;
END_VAR
Filler := CreateFrameworkEvent(Name := Name,
    State := E_State.Idle,
    Severity := E_EventSeverity.Info,
    Message := 'Controlled reservation capacity pressure.');
FOR Index := 1 TO BufferLength DO
    IF FSubject.FreeEntryCount <= FreeCount THEN
        EXIT;
    END_IF;
    IF FSubject.PublishEvent(Event := Filler) <= 0 THEN
        Error(Message := 'Could not create reservation capacity pressure.');
        RETURN;
    END_IF;
END_FOR;
IF FSubject.FreeEntryCount <> FreeCount THEN
    Error(Message := 'Reservation pressure did not reach the intended boundary.');
END_IF;
END_METHOD

{region 'Documentation'}
(*!
<summary>Binds real children, scheduling and isolated storage before introducing capacity pressure.</summary>
*)
{endregion}
METHOD PRIVATE InitializeArrangement
VAR
    Config : ST_TestCaseConfig;
    Index : INT;
END_VAR
IF NOT FSubject.Initialize(Buffer := FEvents,
    FifoControl := FFifo,
    Status := FBufferStatus) THEN
    Error(Message := 'Reservation capture initialization failed.');
    RETURN;
END_IF;
FOwnerReserved := 0;
FOR Index := 1 TO 2 DO
    FChildren[Index].BindPublisher(Publisher := FSubject);
    FChildren[Index].ClearRequestTrace();
    FChildren[Index].ExecutionSlot := INT_TO_UINT(Index);
    IF NOT FChildren[Index].Initialize(Parent := FSubjectParent,
        TestName := CONCAT('AdmissionChild', INT_TO_STRING(Index)),
        Config := Config) THEN
        Error(Message := 'Reservation child initialization failed.');
        RETURN;
    END_IF;
    FChildViews[Index] := FChildren[Index];
    FChildren[Index]();
END_FOR;
IF NOT FCollection.Initialize(Count := 2,
    Children := FChildViews) THEN
    Error(Message := 'Reservation collection initialization failed.');
    RETURN;
END_IF;
FOrchestrator.BindPublisher(Publisher := FSubject);
IF NOT FOrchestrator.Initialize(Collection := FCollection,
    Name := Name) THEN
    Error(Message := 'Reservation Orchestrator initialization failed.');
    RETURN;
END_IF;
SetOwnerReservation(EntryCount := GVL_Constants.TestSuiteResetEventCount,
    Headroom := Param_EventBuffer.EventBufferResetHeadroom);
FillToFreeCount(FreeCount := FOwnerReserved + GVL_Constants.TestCaseResetEventCount
    + Param_EventBuffer.EventBufferResetHeadroom - 1);
FWaitCalls := 0;
FWaitingSequence := FBufferStatus.SequenceId;
END_METHOD

{region 'Documentation'}
(*!
<summary>Completes abort without asynchronous work.</summary>
*)
{endregion}
METHOD PROTECTED ProcessAbort
VAR_INPUT
    Enable : BOOL; //! Phase permission supplied by the owning Test Case; FALSE does not authorize progression, while observation may continue.
END_VAR
IF Enable THEN
    CompleteAbort();
END_IF;
END_METHOD

{region 'Documentation'}
(*!
<summary>Evaluates captured observations after the scenario has finished.</summary>
*)
{endregion}
METHOD PROTECTED ProcessAssertions
VAR_INPUT
    Enable : BOOL; //! Phase permission supplied by the owning Test Case; FALSE does not authorize progression, while observation may continue.
END_VAR
VAR
    Evaluate : BOOL;
END_VAR
Evaluate := Enable AND FPerformed;
FResetWaiting(Enable := Evaluate,
    State := State,
    IN := FResetWaitingMatches);
FExecutionWaiting(Enable := Evaluate,
    State := State,
    IN := FExecutionWaitingMatches);
FReservationBeforeRequest(Enable := Evaluate,
    State := State,
    IN := FReservationBeforeRequestMatches);
FSingleDispatch(Enable := Evaluate,
    State := State,
    IN := FSingleDispatchMatches);
FResumedExecution(Enable := Evaluate,
    State := State,
    IN := FResumedExecutionMatches);
FAccounting(Enable := Evaluate,
    State := State,
    IN := FAccountingMatches);
FConsumerRelease(Enable := Evaluate,
    State := State,
    IN := FConsumerReleaseMatches);
FStorageIntegrity(Enable := Evaluate,
    State := State,
    IN := FStorageIntegrityMatches);
IF Evaluate THEN
    FChecked := TRUE;
END_IF;
END_METHOD

{region 'Documentation'}
(*!
<summary>No Preparation phase is needed.</summary>
*)
{endregion}
METHOD PROTECTED ProcessPreparations
VAR_INPUT
    // SA0033: Required override without Preparation work.
    {attribute 'analysis' := '-33'}
    Enable : BOOL; //! Phase permission supplied by the owning Test Case; FALSE does not authorize progression, while observation may continue.
END_VAR
END_METHOD

{region 'Documentation'}
(*!
<summary>Clears observations; the next attempt initializes fresh isolated storage and child state.</summary>
*)
{endregion}
METHOD PROTECTED ProcessReset
FStep := Setup;
FWaitCalls := 0;
FPerformed := FALSE;
FChecked := FALSE;
FResetWaiting.Reset();
FResetWaitingMatches := TRUE;
FExecutionWaiting.Reset();
FExecutionWaitingMatches := TRUE;
FReservationBeforeRequest.Reset();
FReservationBeforeRequestMatches := TRUE;
FSingleDispatch.Reset();
FSingleDispatchMatches := TRUE;
FResumedExecution.Reset();
FResumedExecutionMatches := TRUE;
FAccounting.Reset();
FAccountingMatches := TRUE;
FConsumerRelease.Reset();
FConsumerReleaseMatches := TRUE;
FStorageIntegrity.Reset();
FStorageIntegrityMatches := TRUE;
FResumedExecutionMatches := FALSE;
CompleteReset();
END_METHOD

{region 'Documentation'}
(*!
<summary>Runs at most one helper/child cycle and waits for final Assertion evaluation.</summary>
*)
{endregion}
METHOD PROTECTED ProcessTests
VAR_INPUT
    Enable : BOOL; //! Phase permission supplied by the owning Test Case; FALSE does not authorize progression, while observation may continue.
END_VAR
IF NOT Enable THEN
    RETURN;
END_IF;
IF FChecked THEN
    CompleteTests();
    RETURN;
END_IF;
IF NOT FPerformed THEN
    RunScenario();
END_IF;
END_METHOD

{region 'Documentation'}
(*!
<summary>Runs the bounded per-cycle admission scenario.</summary>
*)
{endregion}
METHOD PRIVATE RunScenario
CASE FStep OF
    Setup:
        InitializeArrangement();
        IF IsTestingActive THEN
            FStep := WaitForResetCapacity;
        END_IF;

    WaitForResetCapacity:
        CallSubject(Task := E_OrchestratorTask.Reset);
        FResetWaitingMatches := FResetWaitingMatches
            AND (FChildren[1].State = E_State.Uninitialized)
            AND (FChildren[2].State = E_State.Uninitialized)
            AND (FChildren[1].ResetRequestCount = 0)
            AND (FChildren[2].ResetRequestCount = 0)
            AND (FChildren[1].ReservedEntryCount = 0)
            AND (FChildren[2].ReservedEntryCount = 0)
            AND (FBufferStatus.SequenceId = FWaitingSequence);
        FWaitCalls := FWaitCalls + 1;
        IF FWaitCalls = WaitingCalls THEN
            DeletePublishedEvents();
            FStep := CompleteSubjectReset;
        END_IF;

    CompleteSubjectReset:
        CallSubject(Task := E_OrchestratorTask.Reset);
        IF FOrchestrator.IsResetFinished THEN
            FResetWaitingMatches := FResetWaitingMatches
                AND FChildren[1].IsReady AND FChildren[2].IsReady
                AND (FChildren[1].ResetRequestCount = 1)
                AND (FChildren[2].ResetRequestCount = 1);
            FAccountingMatches := FAccountingMatches
                AND (FChildren[1].ReservedEntryCount = 0)
                AND (FChildren[2].ReservedEntryCount = 0);
            FStep := PrepareExecution;
        END_IF;

    PrepareExecution:
        CallSubject(Task := E_OrchestratorTask.Idle);
        IF NOT FOrchestrator.IsReady THEN
            Error(Message := 'Reservation admission arrangement did not become ready.');
            RETURN;
        END_IF;
        DeletePublishedEvents();
        SetOwnerReservation(EntryCount := GVL_Constants.TestSuiteExecutionEventCount,
            Headroom := Param_EventBuffer.EventBufferExecutionHeadroom);
        FillToFreeCount(FreeCount := FOwnerReserved + ChildExecutionBudget
            + Param_EventBuffer.EventBufferExecutionHeadroom - 1);
        FWaitCalls := 0;
        FWaitingSequence := FBufferStatus.SequenceId;
        FStep := WaitForExecutionCapacity;

    WaitForExecutionCapacity:
        CallSubject(Task := E_OrchestratorTask.Execution);
        FExecutionWaitingMatches := FExecutionWaitingMatches
            AND FChildren[1].IsIdle AND FChildren[1].IsReady
            AND FChildren[2].IsIdle AND FChildren[2].IsReady
            AND (FChildren[1].StartRequestCount = 0)
            AND (FChildren[2].StartRequestCount = 0)
            AND (FChildren[1].ReservedEntryCount = 0)
            AND (FChildren[2].ReservedEntryCount = 0)
            AND (FBufferStatus.SequenceId = FWaitingSequence);
        FWaitCalls := FWaitCalls + 1;
        IF FWaitCalls = WaitingCalls THEN
            DeletePublishedEvents();
            FStep := CompleteSubjectExecution;
        END_IF;

    CompleteSubjectExecution:
        CallSubject(Task := E_OrchestratorTask.Execution);
        IF FOrchestrator.IsExecutionFinished THEN
            FResumedExecutionMatches := FChildren[1].IsComplete
                AND FChildren[2].IsComplete
                AND (FChildren[1].Result = E_Result.Passed)
                AND (FChildren[2].Result = E_Result.Passed)
                AND (FChildren[1].StartRequestCount = 1)
                AND (FChildren[2].StartRequestCount = 1);
            FAccountingMatches := FAccountingMatches
                AND (FChildren[1].ReservedEntryCount = 0)
                AND (FChildren[2].ReservedEntryCount = 0);
            FWaitCalls := 0;
            FStep := Finish;
        END_IF;

    Finish:
        CallSubject(Task := E_OrchestratorTask.Execution);
        FWaitCalls := FWaitCalls + 1;
        IF FWaitCalls = WaitingCalls THEN
            SetOwnerReservation(EntryCount := 0,
                Headroom := 0);
            FAccountingMatches := FAccountingMatches AND (FSubject.ReservedEntryCount = 0);
            FPerformed := TRUE;
        END_IF;
ELSE
    Error(Message := 'Unknown reservation admission test step.');
END_CASE;
END_METHOD

{region 'Documentation'}
(*!
<summary>Provides only the concurrent Suite contribution; Suite owner lifecycle is outside this arrangement.</summary>
*)
{endregion}
METHOD PRIVATE SetOwnerReservation
VAR_INPUT
    EntryCount : UINT; //! Replacement concurrent owner reservation after releasing its previous contribution.
    Headroom : UINT; //! Additional free capacity required when reserving the replacement owner contribution.
END_VAR
IF NOT FSubject.FreeReservedSpace(EntryCount := FOwnerReserved,
    OwnerReservedEntryCount := FOwnerReserved) THEN
    Error(Message := 'Concurrent owner reservation release failed.');
    RETURN;
END_IF;
IF NOT FSubject.ReserveSpace(EntryCount := EntryCount,
    HeadroomEntryCount := Headroom,
    OwnerReservedEntryCount := FOwnerReserved) THEN
    Error(Message := 'Concurrent owner reservation failed.');
END_IF;
END_METHOD

END_FUNCTION_BLOCK

// ---- SelfTests/TestCases/TestSuite_EventReservation/Helper/ReservationChildProbe.TcPOU
{region 'Documentation'}
(*!
<summary>Observes reservation state at request entry on a real minimal Test Case.</summary>
<description>
Inherits the normal lifecycle and one real Assertion from SuiteIntegrationChild.
Request overrides only count and observe before delegating to the production method.
No reservation result, state, readiness or scheduling decision is simulated.
ClearRequestTrace clears evidence only, before the isolated scenario begins.
</description>
*)
{endregion}
FUNCTION_BLOCK ReservationChildProbe EXTENDS SuiteIntegrationChild
VAR
    FResetRequestCount : UINT;
    FStartRequestCount : UINT;
    FRequestsReserved : BOOL := TRUE;
END_VAR
VAR CONSTANT
    ExecutionBudget : UINT := 11;
END_VAR

SUPER^();

{region 'Documentation'}
(*!
<summary>Clears observations without changing production lifecycle state.</summary>
*)
{endregion}
METHOD PUBLIC ClearRequestTrace
FResetRequestCount := 0;
FStartRequestCount := 0;
FRequestsReserved := TRUE;
END_METHOD

{region 'Documentation'}
(*!
<summary>Observes the held Reset budget before delegating the request.</summary>
*)
{endregion}
METHOD PUBLIC RequestReset
FResetRequestCount := FResetRequestCount + 1;
FRequestsReserved := FRequestsReserved
    AND (ReservedEntryCount = GVL_Constants.TestCaseResetEventCount)
    AND (EventPublisher.ReservedEntryCount >= ReservedEntryCount);
SUPER^.RequestReset();
END_METHOD

{region 'Documentation'}
(*!
<summary>Retained request-entry observation for the isolated scenario.</summary>
*)
{endregion}
{attribute 'monitoring' := 'call'}
PROPERTY PUBLIC RequestsReserved : BOOL //! Retained request-entry observation for the isolated scenario.
GET
RequestsReserved := FRequestsReserved;
END_GET
END_PROPERTY

{region 'Documentation'}
(*!
<summary>Observes the complete single-Assertion execution budget before delegating.</summary>
*)
{endregion}
METHOD PUBLIC RequestStart
FStartRequestCount := FStartRequestCount + 1;
FRequestsReserved := FRequestsReserved
    AND (ReservedEntryCount = ExecutionBudget)
    AND (EventPublisher.ReservedEntryCount >= ReservedEntryCount);
SUPER^.RequestStart();
END_METHOD

{region 'Documentation'}
(*!
<summary>Retained request-entry observation for the isolated scenario.</summary>
*)
{endregion}
{attribute 'monitoring' := 'call'}
PROPERTY PUBLIC ResetRequestCount : UINT //! Retained request-entry observation for the isolated scenario.
GET
ResetRequestCount := FResetRequestCount;
END_GET
END_PROPERTY

{region 'Documentation'}
(*!
<summary>Retained request-entry observation for the isolated scenario.</summary>
*)
{endregion}
{attribute 'monitoring' := 'call'}
PROPERTY PUBLIC StartRequestCount : UINT //! Retained request-entry observation for the isolated scenario.
GET
StartRequestCount := FStartRequestCount;
END_GET
END_PROPERTY

END_FUNCTION_BLOCK

// ---- SelfTests/TestCases/TestSuite_EventReservation/Test_ImpossibleResetBudget.TcPOU
{region 'Documentation'}
(*!
<summary>Checks an individually impossible reset budget against actual usable capacity.</summary>
<description>

Real subject boundaries

The real Test Case computes reservations; the real Orchestrator decides and publishes its diagnostic.
A collection double supplies one fixed child view. Only the concurrent Suite allowance is held by
the fixture, without running a Suite. Request-entry observations are inherited from the thin child adapter.
The physical array includes one unused FIFO position, leaving capacity one entry below the minimum.
The buffer is empty at rejection: consumer deletion cannot repair an impossible budget.
Three later helper calls must retain Error without another diagnostic or unexpected dispatch.
Expected diagnostics stay in local capture. The surrounding Assertions use the normal selftest publisher.
The real subject binds only local storage; expected findings remain in that storage.
Checking Assertions retain the outer selftest publisher. Each run reinitializes the subject.
</description>
*)
{endregion}
FUNCTION_BLOCK Test_ImpossibleResetBudget EXTENDS TestCaseBase
VAR
    FSubject : EventBuffer;
    FEvents : ARRAY[1..BufferLength] OF ST_Event;
    FFifo : ST_FifoStatus;
    FBufferStatus : ST_EventBufferStatus;
    FPerformed : BOOL;
    FChecked : BOOL;
    FSubjectParent : I_TestSuite;
    FChild : ReservationChildProbe;
    FOrchestrator : OrchestratorProbe;
    FCollection : OrchestrationCollectionDouble;
    FChildren : ARRAY[1..1] OF I_Orchestratable;
    FOwnerReserved : UINT;
    FStep : INT;
    FObservationCalls : UINT;
    FPrecondition : AssertTrue;
    FPreconditionMatches : BOOL;
    FFailureDetection : AssertTrue;
    FFailureDetectionMatches : BOOL;
    FStateAndCounts : AssertTrue;
    FStateAndCountsMatches : BOOL;
    FHeldError : AssertTrue;
    FHeldErrorMatches : BOOL;
    FSingleDiagnostic : AssertTrue;
    FSingleDiagnosticMatches : BOOL;
    FRequestBoundary : AssertTrue;
    FRequestBoundaryMatches : BOOL;
    FAccounting : AssertTrue;
    FAccountingMatches : BOOL;
    FCaptureIntegrity : AssertTrue;
    FCaptureIntegrityMatches : BOOL;
END_VAR
VAR CONSTANT
    BufferLength : UINT := GVL_Constants.TestSuiteResetEventCount + GVL_Constants.TestCaseResetEventCount + Param_EventBuffer.EventBufferResetHeadroom;
    ObservationCalls : UINT := 3;
    ExpectedResetRequests : UINT := 0;
    ExpectedStartRequests : UINT := 0;
    Setup : INT := 0;
    TriggerFailure : INT := 2;
    ObserveFailure : INT := 3;
END_VAR

SUPER^();

{region 'Documentation'}
(*!
<summary>Contributes each checking Assertion once.</summary>
*)
{endregion}
METHOD PROTECTED AggregateResults
VAR_INPUT
    Aggregator : I_ResultAggregator; //! Borrowed result sink owned by the outer Test Case; add this test's checking Assertions without resetting or retaining the sink.
END_VAR
Aggregator.AddProvider(Provider := FPrecondition);
Aggregator.AddProvider(Provider := FFailureDetection);
Aggregator.AddProvider(Provider := FStateAndCounts);
Aggregator.AddProvider(Provider := FHeldError);
Aggregator.AddProvider(Provider := FSingleDiagnostic);
Aggregator.AddProvider(Provider := FRequestBoundary);
Aggregator.AddProvider(Provider := FAccounting);
Aggregator.AddProvider(Provider := FCaptureIntegrity);
END_METHOD

{region 'Documentation'}
(*!
<summary>Supplies only the child identity before initialization.</summary>
*)
{endregion}
METHOD PUBLIC BindSubjectParent
VAR_INPUT
    Parent : I_TestSuite; //! Borrowed identity parent retained for isolated subject initialization; keep the Suite alive through subject use.
END_VAR
FSubjectParent := Parent;
END_METHOD

{region 'Documentation'}
(*!
<summary>Calls the real helper and child and retains accounting observations.</summary>
*)
{endregion}
METHOD PRIVATE CallSubject
VAR_INPUT
    Task : E_OrchestratorTask; //! Orchestration task assigned for this controlled subject call.
END_VAR
FOrchestrator(Task := Task);
FAccountingMatches := FAccountingMatches
    AND (FSubject.ReservedEntryCount = FOwnerReserved + FChild.ReservedEntryCount);
FChild();
FCaptureIntegrityMatches := FCaptureIntegrityMatches
    AND NOT FFifo.ConfigError AND NOT FFifo.IndexError
    AND (FBufferStatus.LostEventCount = 0)
    AND NOT FCollection.InvalidAccess AND NOT FCollection.TraceOverflow;
END_METHOD

{region 'Documentation'}
(*!
<summary>Checks the single retained Orchestrator Error and exact dispatch counts.</summary>
*)
{endregion}
METHOD PRIVATE CheckDiagnostic
VAR
    Index : UINT;
    ErrorCount : UINT;
    PayloadMatches : BOOL := TRUE;
END_VAR
FOR Index := 1 TO BufferLength DO
    IF (FEvents[Index].SequenceId > 0) AND (FEvents[Index].Severity = E_EventSeverity.Error) THEN
        ErrorCount := ErrorCount + 1;
        PayloadMatches := PayloadMatches
            AND (FEvents[Index].OwnerScope = E_OwnerScope.Framework)
            AND (FEvents[Index].EventType = E_EventType.Framework)
            AND (FEvents[Index].State = E_State.Error)
            AND (FEvents[Index].Name = CONCAT(Name, '.Orchestrator'))
            AND (FEvents[Index].Message <> '');
    END_IF;
END_FOR;
FSingleDiagnosticMatches := (ErrorCount = 1) AND PayloadMatches;
FRequestBoundaryMatches := FChild.RequestsReserved
    AND (FChild.ResetRequestCount = ExpectedResetRequests)
    AND (FChild.StartRequestCount = ExpectedStartRequests);
END_METHOD

{region 'Documentation'}
(*!
<summary>Requires all checking Assertions to be initialized.</summary>
*)
{endregion}
METHOD PROTECTED CheckInitialization : BOOL //! TRUE when the inherited initialization check and this concrete fixture check both accept the setup.
CheckInitialization := FALSE;
IF NOT SUPER^.CheckInitialization() OR (FSubjectParent = 0) THEN
    RETURN;
END_IF;

CheckInitialization := FPrecondition.IsInitialized
    AND FFailureDetection.IsInitialized
    AND FStateAndCounts.IsInitialized
    AND FHeldError.IsInitialized
    AND FSingleDiagnostic.IsInitialized
    AND FRequestBoundary.IsInitialized
    AND FAccounting.IsInitialized
    AND FCaptureIntegrity.IsInitialized;
END_METHOD

{region 'Documentation'}
(*!
<summary>Initializes the checking Assertions for one test state.</summary>
*)
{endregion}
METHOD PROTECTED Configure
FPreparationStateCount := 0;
FTestStateCount := 1;
FPrecondition.Initialize(Parent := THIS^,
    AssertionName := 'Precondition');
FFailureDetection.Initialize(Parent := THIS^,
    AssertionName := 'FailureDetection');
FStateAndCounts.Initialize(Parent := THIS^,
    AssertionName := 'StateAndCounts');
FHeldError.Initialize(Parent := THIS^,
    AssertionName := 'HeldError');
FSingleDiagnostic.Initialize(Parent := THIS^,
    AssertionName := 'SingleDiagnostic');
FRequestBoundary.Initialize(Parent := THIS^,
    AssertionName := 'RequestBoundary');
FAccounting.Initialize(Parent := THIS^,
    AssertionName := 'Accounting');
FCaptureIntegrity.Initialize(Parent := THIS^,
    AssertionName := 'CaptureIntegrity');
END_METHOD

{region 'Documentation'}
(*!
<summary>Binds a real child and Orchestrator to fixed isolated storage.</summary>
*)
{endregion}
METHOD PRIVATE InitializeArrangement
VAR
    Config : ST_TestCaseConfig;
END_VAR
IF NOT FSubject.Initialize(Buffer := FEvents,
    FifoControl := FFifo,
    Status := FBufferStatus) THEN
    Error(Message := 'Reservation error capture initialization failed.');
    RETURN;
END_IF;
FOwnerReserved := 0;
FChild.BindPublisher(Publisher := FSubject);
FChild.ClearRequestTrace();
FChild.ExecutionSlot := 1;
IF NOT FChild.Initialize(Parent := FSubjectParent,
    TestName := 'ResetBudgetChild',
    Config := Config) THEN
    Error(Message := 'Reservation error child initialization failed.');
    RETURN;
END_IF;
FChild();
FChildren[1] := FChild;
IF NOT FCollection.Initialize(Count := 1,
    Children := FChildren) THEN
    Error(Message := 'Reservation error collection initialization failed.');
    RETURN;
END_IF;
FOrchestrator.BindPublisher(Publisher := FSubject);
IF NOT FOrchestrator.Initialize(Collection := FCollection,
    Name := Name) THEN
    Error(Message := 'Reservation error Orchestrator initialization failed.');
    RETURN;
END_IF;
IF NOT FSubject.ReserveSpace(EntryCount := GVL_Constants.TestSuiteResetEventCount,
    HeadroomEntryCount := Param_EventBuffer.EventBufferResetHeadroom,
    OwnerReservedEntryCount := FOwnerReserved) THEN
    Error(Message := 'Reservation error concurrent owner setup failed.');
    RETURN;
END_IF;
FPreconditionMatches := FPreconditionMatches AND FChild.IsInitialized
    AND FFifo.BufferEmpty AND (FSubject.Capacity = BufferLength - 1);
END_METHOD

{region 'Documentation'}
(*!
<summary>Completes abort without asynchronous work.</summary>
*)
{endregion}
METHOD PROTECTED ProcessAbort
VAR_INPUT
    Enable : BOOL; //! Phase permission supplied by the owning Test Case; FALSE does not authorize progression, while observation may continue.
END_VAR
IF Enable THEN
    CompleteAbort();
END_IF;
END_METHOD

{region 'Documentation'}
(*!
<summary>Evaluates captured observations after the scenario has finished.</summary>
*)
{endregion}
METHOD PROTECTED ProcessAssertions
VAR_INPUT
    Enable : BOOL; //! Phase permission supplied by the owning Test Case; FALSE does not authorize progression, while observation may continue.
END_VAR
VAR
    Evaluate : BOOL;
END_VAR
Evaluate := Enable AND FPerformed;
FPrecondition(Enable := Evaluate,
    State := State,
    IN := FPreconditionMatches);
FFailureDetection(Enable := Evaluate,
    State := State,
    IN := FFailureDetectionMatches);
FStateAndCounts(Enable := Evaluate,
    State := State,
    IN := FStateAndCountsMatches);
FHeldError(Enable := Evaluate,
    State := State,
    IN := FHeldErrorMatches);
FSingleDiagnostic(Enable := Evaluate,
    State := State,
    IN := FSingleDiagnosticMatches);
FRequestBoundary(Enable := Evaluate,
    State := State,
    IN := FRequestBoundaryMatches);
FAccounting(Enable := Evaluate,
    State := State,
    IN := FAccountingMatches);
FCaptureIntegrity(Enable := Evaluate,
    State := State,
    IN := FCaptureIntegrityMatches);
IF Evaluate THEN
    FChecked := TRUE;
END_IF;
END_METHOD

{region 'Documentation'}
(*!
<summary>No Preparation phase is needed.</summary>
*)
{endregion}
METHOD PROTECTED ProcessPreparations
VAR_INPUT
    // SA0033: Required override without Preparation work.
    {attribute 'analysis' := '-33'}
    Enable : BOOL; //! Phase permission supplied by the owning Test Case; FALSE does not authorize progression, while observation may continue.
END_VAR
END_METHOD

{region 'Documentation'}
(*!
<summary>Clears scenario evidence; next execution initializes a fresh local arrangement.</summary>
*)
{endregion}
METHOD PROTECTED ProcessReset
FStep := Setup;
FObservationCalls := 0;
FPerformed := FALSE;
FChecked := FALSE;
FPrecondition.Reset();
FPreconditionMatches := TRUE;
FFailureDetection.Reset();
FFailureDetectionMatches := TRUE;
FStateAndCounts.Reset();
FStateAndCountsMatches := TRUE;
FHeldError.Reset();
FHeldErrorMatches := TRUE;
FSingleDiagnostic.Reset();
FSingleDiagnosticMatches := TRUE;
FRequestBoundary.Reset();
FRequestBoundaryMatches := TRUE;
FAccounting.Reset();
FAccountingMatches := TRUE;
FCaptureIntegrity.Reset();
FCaptureIntegrityMatches := TRUE;
FSingleDiagnosticMatches := FALSE;
CompleteReset();
END_METHOD

{region 'Documentation'}
(*!
<summary>Advances one scenario phase before checking final captured observations.</summary>
*)
{endregion}
METHOD PROTECTED ProcessTests
VAR_INPUT
    Enable : BOOL; //! Phase permission supplied by the owning Test Case; FALSE does not authorize progression, while observation may continue.
END_VAR
IF NOT Enable THEN
    RETURN;
END_IF;
IF FChecked THEN
    CompleteTests();
    RETURN;
END_IF;
IF NOT FPerformed THEN
    RunScenario();
END_IF;
END_METHOD

{region 'Documentation'}
(*!
<summary>Runs one bounded scenario phase per active outer call.</summary>
*)
{endregion}
METHOD PRIVATE RunScenario
CASE FStep OF
    Setup:
        InitializeArrangement();
        FStep := TriggerFailure;

    TriggerFailure:
        TriggerSubjectFailure();
        FStep := ObserveFailure;

    ObserveFailure:
        CallSubject(Task := E_OrchestratorTask.Reset);
        FFailureDetectionMatches := FFailureDetectionMatches
            AND (FOrchestrator.Result = E_Result.Error);
        FHeldErrorMatches := FHeldErrorMatches
            AND (FOrchestrator.Result = E_Result.Error)
            AND NOT FOrchestrator.IsExecutionFinished;
        FObservationCalls := FObservationCalls + 1;
        IF FObservationCalls = ObservationCalls THEN
            CheckDiagnostic();
            FAccountingMatches := FAccountingMatches
                AND (FChild.ReservedEntryCount = 0);
            IF NOT FSubject.FreeReservedSpace(EntryCount := FOwnerReserved,
                OwnerReservedEntryCount := FOwnerReserved) THEN
                Error(Message := 'Reservation error fixture cleanup failed.');
                RETURN;
            END_IF;
            FAccountingMatches := FAccountingMatches AND (FSubject.ReservedEntryCount = 0);
            FPerformed := TRUE;
        END_IF;
ELSE
    Error(Message := 'Unknown reservation error test step.');
END_CASE;
END_METHOD

{region 'Documentation'}
(*!
<summary>Classifies the impossible budget on an empty buffer, then exercises real Orchestrator handling.</summary>
*)
{endregion}
METHOD PRIVATE TriggerSubjectFailure
VAR
    ReservationResult : E_EventReservationResult;
    PreviousSequence : UDINT;
    PreviousState : E_State;
END_VAR
PreviousSequence := FBufferStatus.SequenceId;
PreviousState := FChild.State;
ReservationResult := FChild.ReserveResetEvents();
FFailureDetectionMatches := ReservationResult = E_EventReservationResult.Error;
FStateAndCountsMatches := (FChild.State = PreviousState)
    AND (FChild.ReservedEntryCount = 0)
    AND (FSubject.ReservedEntryCount = FOwnerReserved)
    AND (FBufferStatus.SequenceId = PreviousSequence)
    AND FFifo.BufferEmpty;
CallSubject(Task := E_OrchestratorTask.Reset);
FFailureDetectionMatches := FFailureDetectionMatches
    AND (FOrchestrator.Result = E_Result.Error);
END_METHOD

END_FUNCTION_BLOCK

// ---- SelfTests/TestCases/TestSuite_EventReservation/Test_ImpossibleExecutionBudget.TcPOU
{region 'Documentation'}
(*!
<summary>Checks an individually impossible execution budget against actual usable capacity.</summary>
<description>

Real subject boundaries

The real Test Case computes reservations; the real Orchestrator decides and publishes its diagnostic.
A collection double supplies one fixed child view. Only the concurrent Suite allowance is held by
the fixture, without running a Suite. Request-entry observations are inherited from the thin child adapter.
The physical array includes one unused FIFO position, leaving capacity one entry below the minimum.
The buffer is empty at rejection: consumer deletion cannot repair an impossible budget.
Three later helper calls must retain Error without another diagnostic or unexpected dispatch.
Expected diagnostics stay in local capture. The surrounding Assertions use the normal selftest publisher.
The real subject binds only local storage; expected findings remain in that storage.
Checking Assertions retain the outer selftest publisher. Each run reinitializes the subject.
</description>
*)
{endregion}
FUNCTION_BLOCK Test_ImpossibleExecutionBudget EXTENDS TestCaseBase
VAR
    FSubject : EventBuffer;
    FEvents : ARRAY[1..BufferLength] OF ST_Event;
    FFifo : ST_FifoStatus;
    FBufferStatus : ST_EventBufferStatus;
    FPerformed : BOOL;
    FChecked : BOOL;
    FSubjectParent : I_TestSuite;
    FChild : ReservationChildProbe;
    FOrchestrator : OrchestratorProbe;
    FCollection : OrchestrationCollectionDouble;
    FChildren : ARRAY[1..1] OF I_Orchestratable;
    FOwnerReserved : UINT;
    FStep : INT;
    FObservationCalls : UINT;
    FPrecondition : AssertTrue;
    FPreconditionMatches : BOOL;
    FFailureDetection : AssertTrue;
    FFailureDetectionMatches : BOOL;
    FStateAndCounts : AssertTrue;
    FStateAndCountsMatches : BOOL;
    FHeldError : AssertTrue;
    FHeldErrorMatches : BOOL;
    FSingleDiagnostic : AssertTrue;
    FSingleDiagnosticMatches : BOOL;
    FRequestBoundary : AssertTrue;
    FRequestBoundaryMatches : BOOL;
    FAccounting : AssertTrue;
    FAccountingMatches : BOOL;
    FCaptureIntegrity : AssertTrue;
    FCaptureIntegrityMatches : BOOL;
END_VAR
VAR CONSTANT
    ChildExecutionBudget : UINT := 11;
    ConfigureExecution : INT := 4;
    BufferLength : UINT := GVL_Constants.TestSuiteExecutionEventCount + ChildExecutionBudget + Param_EventBuffer.EventBufferExecutionHeadroom;
    ObservationCalls : UINT := 3;
    ExpectedResetRequests : UINT := 1;
    ExpectedStartRequests : UINT := 0;
    Setup : INT := 0;
    PrepareChild : INT := 1;
    TriggerFailure : INT := 2;
    ObserveFailure : INT := 3;
END_VAR

SUPER^();

{region 'Documentation'}
(*!
<summary>Contributes each checking Assertion once.</summary>
*)
{endregion}
METHOD PROTECTED AggregateResults
VAR_INPUT
    Aggregator : I_ResultAggregator; //! Borrowed result sink owned by the outer Test Case; add this test's checking Assertions without resetting or retaining the sink.
END_VAR
Aggregator.AddProvider(Provider := FPrecondition);
Aggregator.AddProvider(Provider := FFailureDetection);
Aggregator.AddProvider(Provider := FStateAndCounts);
Aggregator.AddProvider(Provider := FHeldError);
Aggregator.AddProvider(Provider := FSingleDiagnostic);
Aggregator.AddProvider(Provider := FRequestBoundary);
Aggregator.AddProvider(Provider := FAccounting);
Aggregator.AddProvider(Provider := FCaptureIntegrity);
END_METHOD

{region 'Documentation'}
(*!
<summary>Supplies only the child identity before initialization.</summary>
*)
{endregion}
METHOD PUBLIC BindSubjectParent
VAR_INPUT
    Parent : I_TestSuite; //! Borrowed identity parent retained for isolated subject initialization; keep the Suite alive through subject use.
END_VAR
FSubjectParent := Parent;
END_METHOD

{region 'Documentation'}
(*!
<summary>Calls the real helper and child and retains accounting observations.</summary>
*)
{endregion}
METHOD PRIVATE CallSubject
VAR_INPUT
    Task : E_OrchestratorTask; //! Orchestration task assigned for this controlled subject call.
END_VAR
FOrchestrator(Task := Task);
FAccountingMatches := FAccountingMatches
    AND (FSubject.ReservedEntryCount = FOwnerReserved + FChild.ReservedEntryCount);
FChild();
FCaptureIntegrityMatches := FCaptureIntegrityMatches
    AND NOT FFifo.ConfigError AND NOT FFifo.IndexError
    AND (FBufferStatus.LostEventCount = 0)
    AND NOT FCollection.InvalidAccess AND NOT FCollection.TraceOverflow;
END_METHOD

{region 'Documentation'}
(*!
<summary>Checks the single retained Orchestrator Error and exact dispatch counts.</summary>
*)
{endregion}
METHOD PRIVATE CheckDiagnostic
VAR
    Index : UINT;
    ErrorCount : UINT;
    PayloadMatches : BOOL := TRUE;
END_VAR
FOR Index := 1 TO BufferLength DO
    IF (FEvents[Index].SequenceId > 0) AND (FEvents[Index].Severity = E_EventSeverity.Error) THEN
        ErrorCount := ErrorCount + 1;
        PayloadMatches := PayloadMatches
            AND (FEvents[Index].OwnerScope = E_OwnerScope.Framework)
            AND (FEvents[Index].EventType = E_EventType.Framework)
            AND (FEvents[Index].State = E_State.Error)
            AND (FEvents[Index].Name = CONCAT(Name, '.Orchestrator'))
            AND (FEvents[Index].Message <> '');
    END_IF;
END_FOR;
FSingleDiagnosticMatches := (ErrorCount = 1) AND PayloadMatches;
FRequestBoundaryMatches := FChild.RequestsReserved
    AND (FChild.ResetRequestCount = ExpectedResetRequests)
    AND (FChild.StartRequestCount = ExpectedStartRequests);
END_METHOD

{region 'Documentation'}
(*!
<summary>Requires all checking Assertions to be initialized.</summary>
*)
{endregion}
METHOD PROTECTED CheckInitialization : BOOL //! TRUE when the inherited initialization check and this concrete fixture check both accept the setup.
CheckInitialization := FALSE;
IF NOT SUPER^.CheckInitialization() OR (FSubjectParent = 0) THEN
    RETURN;
END_IF;

CheckInitialization := FPrecondition.IsInitialized
    AND FFailureDetection.IsInitialized
    AND FStateAndCounts.IsInitialized
    AND FHeldError.IsInitialized
    AND FSingleDiagnostic.IsInitialized
    AND FRequestBoundary.IsInitialized
    AND FAccounting.IsInitialized
    AND FCaptureIntegrity.IsInitialized;
END_METHOD

{region 'Documentation'}
(*!
<summary>Initializes the checking Assertions for one test state.</summary>
*)
{endregion}
METHOD PROTECTED Configure
FPreparationStateCount := 0;
FTestStateCount := 1;
FPrecondition.Initialize(Parent := THIS^,
    AssertionName := 'Precondition');
FFailureDetection.Initialize(Parent := THIS^,
    AssertionName := 'FailureDetection');
FStateAndCounts.Initialize(Parent := THIS^,
    AssertionName := 'StateAndCounts');
FHeldError.Initialize(Parent := THIS^,
    AssertionName := 'HeldError');
FSingleDiagnostic.Initialize(Parent := THIS^,
    AssertionName := 'SingleDiagnostic');
FRequestBoundary.Initialize(Parent := THIS^,
    AssertionName := 'RequestBoundary');
FAccounting.Initialize(Parent := THIS^,
    AssertionName := 'Accounting');
FCaptureIntegrity.Initialize(Parent := THIS^,
    AssertionName := 'CaptureIntegrity');
END_METHOD

{region 'Documentation'}
(*!
<summary>Binds a real child and Orchestrator to fixed isolated storage.</summary>
*)
{endregion}
METHOD PRIVATE InitializeArrangement
VAR
    Config : ST_TestCaseConfig;
END_VAR
IF NOT FSubject.Initialize(Buffer := FEvents,
    FifoControl := FFifo,
    Status := FBufferStatus) THEN
    Error(Message := 'Reservation error capture initialization failed.');
    RETURN;
END_IF;
FOwnerReserved := 0;
FChild.BindPublisher(Publisher := FSubject);
FChild.ClearRequestTrace();
FChild.ExecutionSlot := 1;
IF NOT FChild.Initialize(Parent := FSubjectParent,
    TestName := 'ExecutionBudgetChild',
    Config := Config) THEN
    Error(Message := 'Reservation error child initialization failed.');
    RETURN;
END_IF;
FChild();
FChildren[1] := FChild;
IF NOT FCollection.Initialize(Count := 1,
    Children := FChildren) THEN
    Error(Message := 'Reservation error collection initialization failed.');
    RETURN;
END_IF;
FOrchestrator.BindPublisher(Publisher := FSubject);
IF NOT FOrchestrator.Initialize(Collection := FCollection,
    Name := Name) THEN
    Error(Message := 'Reservation error Orchestrator initialization failed.');
    RETURN;
END_IF;
IF NOT FSubject.ReserveSpace(EntryCount := GVL_Constants.TestSuiteResetEventCount,
    HeadroomEntryCount := Param_EventBuffer.EventBufferResetHeadroom,
    OwnerReservedEntryCount := FOwnerReserved) THEN
    Error(Message := 'Reservation error concurrent owner setup failed.');
    RETURN;
END_IF;
FPreconditionMatches := FPreconditionMatches AND FChild.IsInitialized
    AND FFifo.BufferEmpty AND (FSubject.Capacity = BufferLength - 1);
END_METHOD

{region 'Documentation'}
(*!
<summary>Removes setup events and replaces the fixture owner allowance; child configuration remains unchanged.</summary>
*)
{endregion}
METHOD PRIVATE PrepareExecution
VAR
    Watermark : UDINT;
END_VAR
Watermark := FBufferStatus.SequenceId;
FSubject.ProcessDeleteRequest(SequenceId := Watermark);
IF NOT FSubject.FreeReservedSpace(EntryCount := FOwnerReserved,
    OwnerReservedEntryCount := FOwnerReserved) THEN
    Error(Message := 'Could not release Reset fixture allowance.');
    RETURN;
END_IF;
IF NOT FSubject.ReserveSpace(EntryCount := GVL_Constants.TestSuiteExecutionEventCount,
    HeadroomEntryCount := Param_EventBuffer.EventBufferExecutionHeadroom,
    OwnerReservedEntryCount := FOwnerReserved) THEN
    Error(Message := 'Could not reserve execution fixture allowance.');
    RETURN;
END_IF;
FPreconditionMatches := FPreconditionMatches AND FFifo.BufferEmpty
    AND (Watermark = 0) AND (FChild.ReservedEntryCount = 0);
END_METHOD

{region 'Documentation'}
(*!
<summary>Completes abort without asynchronous work.</summary>
*)
{endregion}
METHOD PROTECTED ProcessAbort
VAR_INPUT
    Enable : BOOL; //! Phase permission supplied by the owning Test Case; FALSE does not authorize progression, while observation may continue.
END_VAR
IF Enable THEN
    CompleteAbort();
END_IF;
END_METHOD

{region 'Documentation'}
(*!
<summary>Evaluates captured observations after the scenario has finished.</summary>
*)
{endregion}
METHOD PROTECTED ProcessAssertions
VAR_INPUT
    Enable : BOOL; //! Phase permission supplied by the owning Test Case; FALSE does not authorize progression, while observation may continue.
END_VAR
VAR
    Evaluate : BOOL;
END_VAR
Evaluate := Enable AND FPerformed;
FPrecondition(Enable := Evaluate,
    State := State,
    IN := FPreconditionMatches);
FFailureDetection(Enable := Evaluate,
    State := State,
    IN := FFailureDetectionMatches);
FStateAndCounts(Enable := Evaluate,
    State := State,
    IN := FStateAndCountsMatches);
FHeldError(Enable := Evaluate,
    State := State,
    IN := FHeldErrorMatches);
FSingleDiagnostic(Enable := Evaluate,
    State := State,
    IN := FSingleDiagnosticMatches);
FRequestBoundary(Enable := Evaluate,
    State := State,
    IN := FRequestBoundaryMatches);
FAccounting(Enable := Evaluate,
    State := State,
    IN := FAccountingMatches);
FCaptureIntegrity(Enable := Evaluate,
    State := State,
    IN := FCaptureIntegrityMatches);
IF Evaluate THEN
    FChecked := TRUE;
END_IF;
END_METHOD

{region 'Documentation'}
(*!
<summary>No Preparation phase is needed.</summary>
*)
{endregion}
METHOD PROTECTED ProcessPreparations
VAR_INPUT
    // SA0033: Required override without Preparation work.
    {attribute 'analysis' := '-33'}
    Enable : BOOL; //! Phase permission supplied by the owning Test Case; FALSE does not authorize progression, while observation may continue.
END_VAR
END_METHOD

{region 'Documentation'}
(*!
<summary>Clears scenario evidence; next execution initializes a fresh local arrangement.</summary>
*)
{endregion}
METHOD PROTECTED ProcessReset
FStep := Setup;
FObservationCalls := 0;
FPerformed := FALSE;
FChecked := FALSE;
FPrecondition.Reset();
FPreconditionMatches := TRUE;
FFailureDetection.Reset();
FFailureDetectionMatches := TRUE;
FStateAndCounts.Reset();
FStateAndCountsMatches := TRUE;
FHeldError.Reset();
FHeldErrorMatches := TRUE;
FSingleDiagnostic.Reset();
FSingleDiagnosticMatches := TRUE;
FRequestBoundary.Reset();
FRequestBoundaryMatches := TRUE;
FAccounting.Reset();
FAccountingMatches := TRUE;
FCaptureIntegrity.Reset();
FCaptureIntegrityMatches := TRUE;
FSingleDiagnosticMatches := FALSE;
CompleteReset();
END_METHOD

{region 'Documentation'}
(*!
<summary>Advances one scenario phase before checking final captured observations.</summary>
*)
{endregion}
METHOD PROTECTED ProcessTests
VAR_INPUT
    Enable : BOOL; //! Phase permission supplied by the owning Test Case; FALSE does not authorize progression, while observation may continue.
END_VAR
IF NOT Enable THEN
    RETURN;
END_IF;
IF FChecked THEN
    CompleteTests();
    RETURN;
END_IF;
IF NOT FPerformed THEN
    RunScenario();
END_IF;
END_METHOD

{region 'Documentation'}
(*!
<summary>Runs one bounded scenario phase per active outer call.</summary>
*)
{endregion}
METHOD PRIVATE RunScenario
CASE FStep OF
    Setup:
        InitializeArrangement();
        FStep := PrepareChild;

    PrepareChild:
        CallSubject(Task := E_OrchestratorTask.Reset);
        IF FOrchestrator.Result = E_Result.Error THEN
            Error(Message := 'Reservation error scenario could not reset its child.');
            RETURN;
        END_IF;
        IF FOrchestrator.IsResetFinished THEN
            FPreconditionMatches := FPreconditionMatches AND FChild.IsIdle AND FChild.IsReady;
            FStep := ConfigureExecution;
        END_IF;

    ConfigureExecution:
        CallSubject(Task := E_OrchestratorTask.Idle);
        PrepareExecution();
        FStep := TriggerFailure;

    TriggerFailure:
        TriggerSubjectFailure();
        FStep := ObserveFailure;

    ObserveFailure:
        CallSubject(Task := E_OrchestratorTask.Execution);
        FFailureDetectionMatches := FFailureDetectionMatches
            AND (FOrchestrator.Result = E_Result.Error);
        FHeldErrorMatches := FHeldErrorMatches
            AND (FOrchestrator.Result = E_Result.Error)
            AND NOT FOrchestrator.IsExecutionFinished;
        FObservationCalls := FObservationCalls + 1;
        IF FObservationCalls = ObservationCalls THEN
            CheckDiagnostic();
            FAccountingMatches := FAccountingMatches
                AND (FChild.ReservedEntryCount = 0);
            IF NOT FSubject.FreeReservedSpace(EntryCount := FOwnerReserved,
                OwnerReservedEntryCount := FOwnerReserved) THEN
                Error(Message := 'Reservation error fixture cleanup failed.');
                RETURN;
            END_IF;
            FAccountingMatches := FAccountingMatches AND (FSubject.ReservedEntryCount = 0);
            FPerformed := TRUE;
        END_IF;
ELSE
    Error(Message := 'Unknown reservation error test step.');
END_CASE;
END_METHOD

{region 'Documentation'}
(*!
<summary>Classifies the impossible budget on an empty buffer, then exercises real Orchestrator handling.</summary>
*)
{endregion}
METHOD PRIVATE TriggerSubjectFailure
VAR
    ReservationResult : E_EventReservationResult;
    PreviousSequence : UDINT;
    PreviousState : E_State;
END_VAR
PreviousSequence := FBufferStatus.SequenceId;
PreviousState := FChild.State;
ReservationResult := FChild.ReserveExecutionEvents();
FFailureDetectionMatches := ReservationResult = E_EventReservationResult.Error;
FStateAndCountsMatches := (FChild.State = PreviousState)
    AND (FChild.ReservedEntryCount = 0)
    AND (FSubject.ReservedEntryCount = FOwnerReserved)
    AND (FBufferStatus.SequenceId = PreviousSequence)
    AND FFifo.BufferEmpty;
CallSubject(Task := E_OrchestratorTask.Execution);
FFailureDetectionMatches := FFailureDetectionMatches
    AND (FOrchestrator.Result = E_Result.Error);
END_METHOD

END_FUNCTION_BLOCK

// ---- SelfTests/TestCases/TestSuite_EventReservation/Test_ActiveReservationLoss.TcPOU
{region 'Documentation'}
(*!
<summary>Checks Error detection when an active real Test Case loses its event reservation.</summary>
<description>

Real subject boundaries

